        _sut_A._RunExecutionSubstitute();
        _sut_N._RunExecutionSubstitute();
        _done := TRUE;
        ProbeDoneWhen(_done);
    {endregion}
    {region "T505_OnStateChangeWithRestoreCallInside"}
    eTcoSequenceTests.OnStateChangeWithRestoreCallInside:
        IF NOT _arranged THEN
            _sut_A.SetCyclicMode(); //Set sequencer into the cyclic mode
            _sut_N.SetCyclicMode(); //Set sequencer into the cyclic mode
            _sut_A.SetSequenceAsChecked(); //Set sequence as checked, so no StepID uniqueness is performed on next sequence execution
            _sut_N.SetSequenceAsChecked(); //Set sequence as checked, so no StepID uniqueness is performed on next sequence execution
            _sut_A.SetNumberOfSteps(_totalStepNumber); //Set numberOfSteps to the testing instance
            _sut_N.SetNumberOfSteps(_totalStepNumber); //Set numberOfSteps to the testing instance
            _sut_A.TcoSequencerTest := eTcoSequenceTests.OnStateChangeWithRestoreCallInside;
            _sut_N.TcoSequencerTest := eTcoSequenceTests.OnStateChangeWithRestoreCallInside;
            _sut_A.TotalStepNumber := _totalStepNumber;
            _sut_N.TotalStepNumber := _totalStepNumber;
            _sut_A.FinishStep := FALSE;
            _sut_N.FinishStep := FALSE;
            _plcCycleCounter := 0;
            _arranged := TRUE;
            RETURN;
        END_IF

        IF NOT _done THEN
            IF _plcCycleCounter = 1 THEN
                _sut_A.CallRestoreInOnStateChange := FALSE;
                _sut_N.CallRestoreInOnStateChange := FALSE;
            ELSE
                _sut_A.CallRestoreInOnStateChange := TRUE;
                _sut_N.CallRestoreInOnStateChange := TRUE;
                _sut_A.FinishStep := TRUE;
                _sut_N.FinishStep := TRUE;
            END_IF

            _sut_A._RunExecutionSubstitute();
            _sut_N._RunExecutionSubstitute();
        END_IF

        _done := _plcCycleCounter >= 2;

        IF _done THEN
            _sut_A.CallRestoreInOnStateChange := FALSE;
            _sut_N.CallRestoreInOnStateChange := FALSE;
            ProbeDoneWhen(_done);
        END_IF
    {endregion}
    {region "T506_MinStepId"}
    eTcoSequenceTests.MinStepId:
        IF NOT _arranged THEN
            _sut_A.SetCyclicMode(); //Set sequencer into the cyclic mode
            _sut_N.SetCyclicMode(); //Set sequencer into the cyclic mode
            _sut_A.SetSequenceAsChecked(); //Set sequence as checked, so no StepID uniqueness is performed on next sequence execution
            _sut_N.SetSequenceAsChecked(); //Set sequence as checked, so no StepID uniqueness is performed on next sequence execution
            _sut_A.SetNumberOfSteps(_totalStepNumber); //Set numberOfSteps to the testing instance
            _sut_N.SetNumberOfSteps(_totalStepNumber); //Set numberOfSteps to the testing instance
            _sut_A.TcoSequencerTest := eTcoSequenceTests.MinStepId;
            _sut_N.TcoSequencerTest := eTcoSequenceTests.MinStepId;
            _sut_A.TotalStepNumber := _totalStepNumber;
            _sut_N.TotalStepNumber := _totalStepNumber;
            _sut_A.FinishStep := FALSE;
            _sut_N.FinishStep := FALSE;
            _plcCycleCounter := 0;
            _arranged := TRUE;
            RETURN;
        END_IF

        IF NOT _done THEN
            _sut_A.StepId := _currentStepId;
            _sut_N.StepId := _currentStepId;
            _sut_A._RunExecutionSubstitute();
            _sut_N._RunExecutionSubstitute();
        END_IF

        _done := TRUE;
        ProbeDoneWhen(_done);
    {endregion}
    {region "T507_MaxStepId"}
    eTcoSequenceTests.MaxStepId:
        IF NOT _arranged THEN
            _sut_A.SetCyclicMode(); //Set sequencer into the cyclic mode
            _sut_N.SetCyclicMode(); //Set sequencer into the cyclic mode
            _sut_A.SetSequenceAsChecked(); //Set sequence as checked, so no StepID uniqueness is performed on next sequence execution
            _sut_N.SetSequenceAsChecked(); //Set sequence as checked, so no StepID uniqueness is performed on next sequence execution
            _sut_A.SetNumberOfSteps(_totalStepNumber); //Set numberOfSteps to the testing instance
            _sut_N.SetNumberOfSteps(_totalStepNumber); //Set numberOfSteps to the testing instance
            _sut_A.TcoSequencerTest := eTcoSequenceTests.MaxStepId;
            _sut_N.TcoSequencerTest := eTcoSequenceTests.MaxStepId;
            _sut_A.TotalStepNumber := _totalStepNumber;
            _sut_N.TotalStepNumber := _totalStepNumber;
            _sut_A.FinishStep := FALSE;
            _sut_N.FinishStep := FALSE;
            _plcCycleCounter := 0;
            _arranged := TRUE;
            RETURN;
        END_IF

        IF NOT _done THEN
            _sut_A.StepId := _currentStepId;
            _sut_N.StepId := _currentStepId;
            _sut_A._RunExecutionSubstitute();
            _sut_N._RunExecutionSubstitute();
        END_IF

        _done := TRUE;
        ProbeDoneWhen(_done);
    {endregion}
    {region "T508_RequestStepToFirstStepWithStepId0"}
    eTcoSequenceTests.RequestStepToFirstStepWithStepId0:
        IF NOT _arranged THEN
            _sut_A.SetCyclicMode(); //Set sequencer into the cyclic mode
            _sut_N.SetCyclicMode(); //Set sequencer into the cyclic mode
            _sut_A.SetSequenceAsChecked(); //Set sequence as checked, so no StepID uniqueness is performed on next sequence execution
            _sut_N.SetSequenceAsChecked(); //Set sequence as checked, so no StepID uniqueness is performed on next sequence execution
            _sut_A.SetNumberOfSteps(_totalStepNumber); //Set numberOfSteps to the testing instance
            _sut_N.SetNumberOfSteps(_totalStepNumber); //Set numberOfSteps to the testing instance
            _sut_A.TcoSequencerTest := eTcoSequenceTests.RequestStepToFirstStepWithStepId0;
            _sut_N.TcoSequencerTest := eTcoSequenceTests.RequestStepToFirstStepWithStepId0;
            _sut_A.TotalStepNumber := _totalStepNumber;
            _sut_N.TotalStepNumber := _totalStepNumber;
            _sut_A.FinishStep := TRUE;
            _sut_N.FinishStep := TRUE;
            _plcCycleCounter := 0;
            _arranged := TRUE;
            RETURN;
        END_IF

        IF NOT _done THEN
            IF _plcCycleCounter > 1 THEN
                _sut_A.FinishStep := FALSE;
                _sut_N.FinishStep := FalsE;
            END_IF

            _sut_A._RunExecutionSubstitute();
            _sut_N._RunExecutionSubstitute();
        END_IF

        _done := _plcCycleCounter > 1;
        ProbeDoneWhen(_done);
    {endregion}
    {region "T509_RequestStep"}
    eTcoSequenceTests.RequestStep:
        IF NOT _arranged THEN
            _sut_A.SetCyclicMode(); //Set sequencer into the cyclic mode
            _sut_N.SetCyclicMode(); //Set sequencer into the cyclic mode
            _sut_A.SetSequenceAsChecked(); //Set sequence as checked, so no StepID uniqueness is performed on next sequence execution
            _sut_N.SetSequenceAsChecked(); //Set sequence as checked, so no StepID uniqueness is performed on next sequence execution
            _sut_A.SetNumberOfSteps(10); //Set numberOfSteps to the testing instance
            _sut_N.SetNumberOfSteps(10); //Set numberOfSteps to the testing instance
            _sut_A.TcoSequencerTest := eTcoSequenceTests.RequestStep;
            _sut_N.TcoSequencerTest := eTcoSequenceTests.RequestStep;
            _plcCycleCounter := 0;
            _arranged := TRUE;
            RETURN;
        END_IF

        IF NOT _done THEN
            _sut_A.SequenceRun := _plcCycleCounter;
            _sut_N.SequenceRun := _plcCycleCounter;
            _sut_A._RunExecutionSubstitute();
            _sut_N._RunExecutionSubstitute();
        END_IF

        _done := _plcCycleCounter >= 3;
        ProbeDoneWhen(_done);
    {endregion}
    {region "T510_CheckStepIdUniqueness"}
    eTcoSequenceTests.CheckStepIdUniqueness:
        IF NOT _arranged THEN
            _sut_A.SetCyclicMode(); //Set sequencer into the cyclic mode
            _sut_N.SetCyclicMode(); //Set sequencer into the cyclic mode
            _sut_A.SetSequenceAsNotChecked(); //Set sequence as not checked, so StepId uniqueness is going to be performed on next sequence run
            _sut_N.SetSequenceAsNotChecked(); //Set sequence as not checked, so StepId uniqueness is going to be performed on next sequence run
            _sut_A.ClearNumberOfSteps(); //Clear internal step counters, so number of steps is going to be counted again on next sequence run
            _sut_N.ClearNumberOfSteps(); //Clear internal step counters, so number of steps is going to be counted again on next sequence run
            _sut_A.Enabled := TRUE;
            _sut_A.RunOneStep := FALSE;
            _sut_A.RunAllSteps := TRUE;
            _sut_A.FinishStep := TRUE;
            _sut_N.Enabled := TRUE;
            _sut_N.RunOneStep := FALSE;
            _sut_N.RunAllSteps := TRUE;
            _sut_N.FinishStep := TRUE;
            _sut_A.SetCurrentStep(inStepID := _currentStepId, inStepDescription := _currentStepDescription);
            _sut_N.SetCurrentStep(inStepID := _currentStepId, inStepDescription := _currentStepDescription);
            _sut_A.TcoSequencerTest := eTcoSequenceTests.CheckStepIdUniqueness;
            _sut_N.TcoSequencerTest := eTcoSequenceTests.CheckStepIdUniqueness;
            _sut_A.SaveNumberOfStepsInSequence();
            _sut_N.SaveNumberOfStepsInSequence();
            _plcCycleCounter := 0;
            _arranged := TRUE;
            RETURN;
        END_IF

        IF NOT _done THEN
            _sut_A._RunExecutionSubstitute();
            _sut_N._RunExecutionSubstitute();
            _sut_A.SaveNumberOfStepsInSequence();
            _sut_N.SaveNumberOfStepsInSequence();
        END_IF

        _done := _plcCycleCounter >= 2;
        ProbeDoneWhen(_done);
    {endregion}
    {region "T512_RestoreAlreadyCheckedSequence"}
    eTcoSequenceTests.RestoreAlreadyCheckedSequence:
        _sut_A.Restore();
        _sut_N.Restore();
        _sut_A.SaveNumberOfStepsInSequence();
        _sut_N.SaveNumberOfStepsInSequence();
        _done := TRUE;
        ProbeDoneWhen(_done);
    {endregion}
    {region "T513_CheckStepIdUniqueness"}
    eTcoSequenceTests.NotUniqueStepId:
        IF NOT _arranged THEN
            _sut_A.Enabled := TRUE;
            _sut_A.RunOneStep := FALSE;
            _sut_A.RunAllSteps := FALSE;
            _sut_A.FinishStep := TRUE;
            _sut_A.StepId := _stepId;
            _sut_N.Enabled := TRUE;
            _sut_N.RunOneStep := FALSE;
            _sut_N.RunAllSteps := FALSE;
            _sut_N.FinishStep := TRUE;
            _sut_N.StepId := _stepId;
            _sut_A.SetCurrentStep(inStepID := _currentStepId, inStepDescription := _currentStepDescription);
            _sut_N.SetCurrentStep(inStepID := _currentStepId, inStepDescription := _currentStepDescription);
            _sut_A.TcoSequencerTest := eTcoSequenceTests.NotUniqueStepId;
            _sut_N.TcoSequencerTest := eTcoSequenceTests.NotUniqueStepId;
            _sut_A.SaveNumberOfStepsInSequence();
            _sut_N.SaveNumberOfStepsInSequence();
            _plcCycleCounter := 0;
			_sut_A._messenger.Clear();
			_sut_N._messenger.Clear();
            _arranged := TRUE;
            RETURN;
        END_IF

        IF NOT _done THEN								 
            _sut_A._RunExecutionSubstitute();
            _sut_N._RunExecutionSubstitute();
            _sut_A.SaveNumberOfStepsInSequence();
            _sut_N.SaveNumberOfStepsInSequence();
            _done := _plcCycleCounter >= 2;
        END_IF

        IF _done THEN
            ProbeDoneWhen(_done);
        END_IF
    {endregion}
    {region "T516_AfterErrorRestore"}
    eTcoSequenceTests.AfterErrorRestore:
        IF NOT _arranged THEN
            _sut_A.TcoSequencerTest := eTcoSequenceTests.AfterErrorRestore;
            _sut_N.TcoSequencerTest := eTcoSequenceTests.AfterErrorRestore;
            _sut_A.SaveNumberOfStepsInSequence();
            _sut_N.SaveNumberOfStepsInSequence();
            _plcCycleCounter := 0;
            _arranged := TRUE;
            RETURN;
        END_IF

        IF NOT _done THEN
            _sut_A._RunExecutionSubstitute();
            _sut_N._RunExecutionSubstitute();
            _sut_A.SaveNumberOfStepsInSequence();
            _sut_N.SaveNumberOfStepsInSequence();
            _done := _plcCycleCounter >= 3;
        END_IF

        IF _done THEN
            ProbeDoneWhen(_done);
        END_IF
    {endregion}
    {region "T520_ChangeStepIdDuringExecution"}
    eTcoSequenceTests.ChangeStepIdDuringExecution:
        IF NOT _arranged THEN
            _sut_A.TcoSequencerTest := eTcoSequenceTests.ChangeStepIdDuringExecution;
            _sut_N.TcoSequencerTest := eTcoSequenceTests.ChangeStepIdDuringExecution;
            _sut_A.SetCyclicMode(); //Set sequencer into the cyclic mode
            _sut_N.SetCyclicMode(); //Set sequencer into the cyclic mode
            _sut_A.SetSequenceAsChecked(); //Set sequence as checked, so no StepID uniqueness is performed on next sequence execution
            _sut_N.SetSequenceAsChecked(); //Set sequence as checked, so no StepID uniqueness is performed on next sequence execution
            _sut_A.ClearNumberOfSteps(); //Clear internal step counters, so number of steps is going to be counted again on next sequence run
            _sut_N.ClearNumberOfSteps(); //Clear internal step counters, so number of steps is going to be counted again on next sequence run
            _sut_A.SetCurrentStep(inStepID := _currentStepId, inStepDescription := _currentStepDescription);
            _sut_N.SetCurrentStep(inStepID := _currentStepId, inStepDescription := _currentStepDescription);
            _sut_A.TotalStepNumber := _totalStepNumber;
            _sut_N.TotalStepNumber := _totalStepNumber;
            _sut_A.SaveNumberOfStepsInSequence();
            _sut_N.SaveNumberOfStepsInSequence();
            _plcCycleCounter := 0;
            _arranged := TRUE;
            RETURN;
        END_IF

        IF NOT _done THEN
            _sut_A.SequenceRun := _plcCycleCounter;
            _sut_N.SequenceRun := _plcCycleCounter;
            _sut_A._RunExecutionSubstitute();
            _sut_N._RunExecutionSubstitute();
            _sut_A.SaveNumberOfStepsInSequence();
            _sut_N.SaveNumberOfStepsInSequence();
        END_IF

        _done := _plcCycleCounter >= 3;
        ProbeDoneWhen(_done);
    {endregion}
    {region "T524_CommentOutPartOfRunningSequencer"}
    eTcoSequenceTests.CommentOutPartOfRunningSequencer:
        IF NOT _arranged THEN
            _sut_A.TcoSequencerTest := eTcoSequenceTests.CommentOutPartOfRunningSequencer;
            _sut_N.TcoSequencerTest := eTcoSequenceTests.CommentOutPartOfRunningSequencer;
            _sut_A.SetCyclicMode(); //Set sequencer into the cyclic mode
            _sut_N.SetCyclicMode(); //Set sequencer into the cyclic mode
            _sut_A.SetSequenceAsChecked(); //Set sequence as checked, so no StepID uniqueness is performed on next sequence execution
            _sut_N.SetSequenceAsChecked(); //Set sequence as checked, so no StepID uniqueness is performed on next sequence execution
            _sut_A.ClearNumberOfSteps(); //Clear internal step counters, so number of steps is going to be counted again on next sequence run
            _sut_N.ClearNumberOfSteps(); //Clear internal step counters, so number of steps is going to be counted again on next sequence run
            _sut_A.SetCurrentStep(inStepID := _currentStepId, inStepDescription := _currentStepDescription);
            _sut_N.SetCurrentStep(inStepID := _currentStepId, inStepDescription := _currentStepDescription);
            _sut_A.TotalStepNumber := _totalStepNumber;
            _sut_N.TotalStepNumber := _totalStepNumber;
            _sut_A.SaveNumberOfStepsInSequence();
            _sut_N.SaveNumberOfStepsInSequence();
            _plcCycleCounter := 0;
            _arranged := TRUE;
            RETURN;
        END_IF

        IF NOT _done THEN
            IF _plcCycleCounter = 3 THEN
                _sut_A.Restore();
                _sut_N.Restore();
                _sut_A.SetSequenceAsChecked(); //Set sequence as checked, so no StepID uniqueness is performed on next sequence execution
                _sut_N.SetSequenceAsChecked(); //Set sequence as checked, so no StepID uniqueness is performed on next sequence execution
                _sut_A.ClearNumberOfSteps(); //Clear internal step counters, so number of steps is going to be counted again on next sequence run
                _sut_N.ClearNumberOfSteps(); //Clear internal step counters, so number of steps is going to be counted again on next sequence run
            END_IF

            _sut_A.SequenceRun := _plcCycleCounter;
            _sut_N.SequenceRun := _plcCycleCounter;
            _sut_A._RunExecutionSubstitute();
            _sut_N._RunExecutionSubstitute();
            _sut_A.SaveNumberOfStepsInSequence();
            _sut_N.SaveNumberOfStepsInSequence();
        END_IF

        _done := _plcCycleCounter >= 3;
        ProbeDoneWhen(_done);
    {endregion}
    {region "T526_UncommentPartOfRunningSequencer"}
    eTcoSequenceTests.UncommentPartOfRunningSequencer:
        IF NOT _arranged THEN
            _sut_A.TcoSequencerTest := eTcoSequenceTests.UncommentPartOfRunningSequencer;
            _sut_N.TcoSequencerTest := eTcoSequenceTests.UncommentPartOfRunningSequencer;
            _sut_A.SetCyclicMode(); //Set sequencer into the cyclic mode
            _sut_N.SetCyclicMode(); //Set sequencer into the cyclic mode
            _sut_A.SetSequenceAsChecked(); //Set sequence as checked, so no StepID uniqueness is performed on next sequence execution
            _sut_N.SetSequenceAsChecked(); //Set sequence as checked, so no StepID uniqueness is performed on next sequence execution
            _sut_A.ClearNumberOfSteps(); //Clear internal step counters, so number of steps is going to be counted again on next sequence run
            _sut_N.ClearNumberOfSteps(); //Clear internal step counters, so number of steps is going to be counted again on next sequence run
            _sut_A.SetCurrentStep(inStepID := _currentStepId, inStepDescription := _currentStepDescription);
            _sut_N.SetCurrentStep(inStepID := _currentStepId, inStepDescription := _currentStepDescription);
            _sut_A.TotalStepNumber := _totalStepNumber;
            _sut_N.TotalStepNumber := _totalStepNumber;
            _sut_A.SaveNumberOfStepsInSequence();
            _sut_N.SaveNumberOfStepsInSequence();
            _plcCycleCounter := 0;
            _arranged := TRUE;
            RETURN;
        END_IF

        IF NOT _done THEN
            _sut_A.SequenceRun := _plcCycleCounter;
            _sut_N.SequenceRun := _plcCycleCounter;
            _sut_A._RunExecutionSubstitute();
            _sut_N._RunExecutionSubstitute();
            _sut_A.SaveNumberOfStepsInSequence();
            _sut_N.SaveNumberOfStepsInSequence();
        END_IF

        _done := _plcCycleCounter >= 2;
        ProbeDoneWhen(_done);
    {endregion}
    {region "T530_OpenCloseSequence"}
    eTcoSequenceTests.OpenCloseSequence:
        IF NOT _arranged THEN
            _sut_A.TcoSequencerTest := eTcoSequenceTests.OpenCloseSequence;
            _sut_N.TcoSequencerTest := eTcoSequenceTests.OpenCloseSequence;
            _sut_A.SetCyclicMode(); //Set sequencer into the cyclic mode
            _sut_N.SetCyclicMode(); //Set sequencer into the cyclic mode
            _sut_A.SetSequenceAsChecked(); //Set sequence as checked, so no StepID uniqueness is performed on next sequence execution
            _sut_N.SetSequenceAsChecked(); //Set sequence as checked, so no StepID uniqueness is performed on next sequence execution
            _sut_A.ClearNumberOfSteps(); //Clear internal step counters, so number of steps is going to be counted again on next sequence run
            _sut_N.ClearNumberOfSteps(); //Clear internal step counters, so number of steps is going to be counted again on next sequence run
            _sut_A.TotalStepNumber := _totalStepNumber;
            _sut_N.TotalStepNumber := _totalStepNumber;
            _sut_A.SaveNumberOfStepsInSequence();
            _sut_N.SaveNumberOfStepsInSequence();
            _plcCycleCounter := 0;
            _arranged := TRUE;
            RETURN;
        END_IF

        IF NOT _done THEN
            IF _plcCycleCounter = 1 THEN
                _sut_A.SequencerOpen();
                _sut_N.SequencerOpen();

                IF _sut_A._Step(0, TRUE, 'Step 0') THEN
                    _sut_A._StepCompleteWhen(TRUE);
                END_IF

                IF _sut_N._Step(0, TRUE, 'Step 0') THEN
                    _sut_N._StepCompleteWhen(TRUE);
                END_IF
				_sut_A.SequencerClose();
                _sut_N.SequencerClose();
            END_IF

            IF _plcCycleCounter = 2 THEN
				_sut_A.SequencerOpen();
                _sut_N.SequencerOpen();
                FOR i := 1 TO _totalStepNumber DO
                    _sut_A._Step(i, TRUE, CONCAT('Step ', INT_TO_STRING(i)));
                    _sut_N._Step(i, TRUE, CONCAT('Step ', INT_TO_STRING(i)));
                END_FOR

                _sut_A.SequencerClose();
                _sut_N.SequencerClose();
            END_IF
		END_IF;		 
		
        _done := _plcCycleCounter >= 2;
        ProbeDoneWhen(_done);			  

//            IF _plcCycleCounter = 3 THEN
//                _sut_A.SequencerOpen();
//                _sut_N.SequencerOpen();
//			    _sut_A.SequencerClose();
//                _sut_N.SequencerClose();
//            END_IF

//            IF _plcCycleCounter = 4 THEN
//				_sut_A.SequencerOpen();
//                _sut_N.SequencerOpen();
//                IF _sut_A._Step(0, TRUE, 'Step 0') THEN
//                    _sut_A._StepCompleteWhen(TRUE);
//                END_IF

//                IF _sut_N._Step(0, TRUE, 'Step 0') THEN
//                    _sut_N._StepCompleteWhen(TRUE);
//                END_IF
//				_sut_A.SequencerClose();
//                _sut_N.SequencerClose();	 
//            END_IF

//            IF _plcCycleCounter = 5 THEN
//				_sut_A.SequencerOpen();
//                _sut_N.SequencerOpen();
//                FOR i := 1 TO _totalStepNumber DO
//                    IF _sut_A._Step(i, TRUE, CONCAT('Step ', INT_TO_STRING(i))) THEN
//                        _sut_A._StepCompleteWhen(TRUE);
//                    END_IF

//                    IF _sut_N._Step(i, TRUE, CONCAT('Step ', INT_TO_STRING(i))) THEN
//                        _sut_N._StepCompleteWhen(TRUE);
//                    END_IF
//                END_FOR
//				_sut_A.SequencerClose();
//                _sut_N.SequencerClose();	 
//            END_IF

//            IF _plcCycleCounter = 6 THEN
//                _sut_A._SequenceComplete();
//                _sut_N._SequenceComplete();
//                _sut_A.SequencerClose();
//                _sut_N.SequencerClose();
//            END_IF

//            IF _plcCycleCounter = 7 THEN
//                _sut_A.SequencerOpen();
//                _sut_N.SequencerOpen();
//            END_IF

//            IF _plcCycleCounter = 8 THEN
//                _sut_A.SequencerClose();
//                _sut_N.SequencerClose();
//            END_IF

//            IF _plcCycleCounter = 9 THEN
//                _sut_A.SequencerOpen();
//                _sut_N.SequencerOpen();
//                _sut_A._Step(0, TRUE, 'Step 0');
//                _sut_N._Step(0, TRUE, 'Step 0');
//                _sut_A.SequencerClose();
//                _sut_N.SequencerClose();
//            END_IF
//        END_IF

//        _done := _plcCycleCounter >= 9;
//        ProbeDoneWhen(_done);
    {endregion}
    {region "T541_RequestStepFromLowerToHigher"}
    eTcoSequenceTests.RequestStepFromLowerToHigher:
        IF NOT _arranged THEN
            _sut_A.TcoSequencerTest := eTcoSequenceTests.RequestStepFromLowerToHigher;
            _sut_N.TcoSequencerTest := eTcoSequenceTests.RequestStepFromLowerToHigher;
            _sut_A.SetCyclicMode(); //Set sequencer into the cyclic mode
            _sut_N.SetCyclicMode(); //Set sequencer into the cyclic mode
            _sut_A.SetSequenceAsChecked(); //Set sequence as checked, so no StepID uniqueness is performed on next sequence execution
            _sut_N.SetSequenceAsChecked(); //Set sequence as checked, so no StepID uniqueness is performed on next sequence execution
            _sut_A.ClearNumberOfSteps(); //Clear internal step counters, so number of steps is going to be counted again on next sequence run
            _sut_N.ClearNumberOfSteps(); //Clear internal step counters, so number of steps is going to be counted again on next sequence run
            _sut_A.SetCurrentStep(inStepID := _currentStepId, inStepDescription := _currentStepDescription);
            _sut_N.SetCurrentStep(inStepID := _currentStepId, inStepDescription := _currentStepDescription);
            _sut_A.TotalStepNumber := _totalStepNumber;
            _sut_N.TotalStepNumber := _totalStepNumber;
            _sut_A.ReqStep := _reqStep;
            _sut_N.ReqStep := _reqStep;
            _sut_A.ReqStepNotExists := _reqStepNotExists;
            _sut_N.ReqStepNotExists := _reqStepNotExists;
            _sut_A.SaveNumberOfStepsInSequence();
            _sut_N.SaveNumberOfStepsInSequence();
            _plcCycleCounter := 0;
            _arranged := TRUE;
            RETURN;
        END_IF

        IF NOT _done THEN
            _sut_A.SequenceRun := _plcCycleCounter;
            _sut_N.SequenceRun := _plcCycleCounter;
            _sut_A._RunExecutionSubstitute();
            _sut_N._RunExecutionSubstitute();
            _sut_A.SaveNumberOfStepsInSequence();
            _sut_N.SaveNumberOfStepsInSequence();
        END_IF

        _done := _plcCycleCounter >= 2;
        ProbeDoneWhen(_done);
    {endregion}
    {region "T542_RequestStepFromHigherToLower"}
    eTcoSequenceTests.RequestStepFromHigherToLower:
        IF NOT _arranged THEN
            _sut_A.TcoSequencerTest := eTcoSequenceTests.RequestStepFromHigherToLower;
            _sut_N.TcoSequencerTest := eTcoSequenceTests.RequestStepFromHigherToLower;
            _sut_A.SetCyclicMode(); //Set sequencer into the cyclic mode
            _sut_N.SetCyclicMode(); //Set sequencer into the cyclic mode
            _sut_A.SetSequenceAsChecked(); //Set sequence as checked, so no StepID uniqueness is performed on next sequence execution
            _sut_N.SetSequenceAsChecked(); //Set sequence as checked, so no StepID uniqueness is performed on next sequence execution
            _sut_A.SetNumberOfSteps(_totalStepNumber);
            _sut_N.SetNumberOfSteps(_totalStepNumber);
            _sut_A.SetCurrentStep(inStepID := _currentStepId, inStepDescription := _currentStepDescription);
            _sut_N.SetCurrentStep(inStepID := _currentStepId, inStepDescription := _currentStepDescription);
            _sut_A.TotalStepNumber := _totalStepNumber;
            _sut_N.TotalStepNumber := _totalStepNumber;
            _sut_A.ReqStep := _reqStep;
            _sut_N.ReqStep := _reqStep;
            _sut_A.ReqStepNotExists := _reqStepNotExists;
            _sut_N.ReqStepNotExists := _reqStepNotExists;
            _sut_A.SaveNumberOfStepsInSequence();
            _sut_N.SaveNumberOfStepsInSequence();
            _plcCycleCounter := 0;
            _arranged := TRUE;
            RETURN;
        END_IF

        IF NOT _done THEN
            _sut_A.SequenceRun := _plcCycleCounter;
            _sut_N.SequenceRun := _plcCycleCounter;
            _sut_A._RunExecutionSubstitute();
            _sut_N._RunExecutionSubstitute();
            _sut_A.SaveNumberOfStepsInSequence();
            _sut_N.SaveNumberOfStepsInSequence();
        END_IF

        _done := _plcCycleCounter >= 2;
        ProbeDoneWhen(_done);
    {endregion}
    {region "T544_RequestStepToNotExistingStep"}
    eTcoSequenceTests.RequestStepToNotExistingStep:
        IF NOT _arranged THEN
            _sut_A.TcoSequencerTest := eTcoSequenceTests.RequestStepToNotExistingStep;
            _sut_N.TcoSequencerTest := eTcoSequenceTests.RequestStepToNotExistingStep;
            _sut_A.SetCyclicMode(); //Set sequencer into the cyclic mode
            _sut_N.SetCyclicMode(); //Set sequencer into the cyclic mode
            _sut_A.SetSequenceAsChecked(); //Set sequence as checked, so no StepID uniqueness is performed on next sequence execution
            _sut_N.SetSequenceAsChecked(); //Set sequence as checked, so no StepID uniqueness is performed on next sequence execution
            _sut_A.SetNumberOfSteps(_totalStepNumber);
            _sut_N.SetNumberOfSteps(_totalStepNumber);
            _sut_A.SetCurrentStep(inStepID := _currentStepId, inStepDescription := _currentStepDescription);
            _sut_N.SetCurrentStep(inStepID := _currentStepId, inStepDescription := _currentStepDescription);
            _sut_A.TotalStepNumber := _totalStepNumber;
            _sut_N.TotalStepNumber := _totalStepNumber;
            _sut_A.ReqStep := _reqStep;
            _sut_N.ReqStep := _reqStep;
            _sut_A.ReqStepNotExists := _reqStepNotExists;
            _sut_N.ReqStepNotExists := _reqStepNotExists;
            _sut_A.SaveNumberOfStepsInSequence();
            _sut_N.SaveNumberOfStepsInSequence();
            _plcCycleCounter := 0;
            _arranged := TRUE;
            RETURN;
        END_IF

        IF _plcCycleCounter = 4 THEN
            _sut_A.Restore();
            _sut_N.Restore();
            _sut_A.SetCyclicMode(); //Set sequencer into the cyclic mode
            _sut_N.SetCyclicMode(); //Set sequencer into the cyclic mode
            _sut_A.SetSequenceAsChecked(); //Set sequence as checked, so no StepID uniqueness is performed on next sequence execution
            _sut_N.SetSequenceAsChecked(); //Set sequence as checked, so no StepID uniqueness is performed on next sequence execution
            _sut_A.SetNumberOfSteps(_totalStepNumber);
            _sut_N.SetNumberOfSteps(_totalStepNumber);
            _sut_A.SetCurrentStep(inStepID := _currentStepId, inStepDescription := _currentStepDescription);
            _sut_N.SetCurrentStep(inStepID := _currentStepId, inStepDescription := _currentStepDescription);
            _sut_A.TotalStepNumber := _totalStepNumber;
            _sut_N.TotalStepNumber := _totalStepNumber;
        END_IF

        IF NOT _done THEN
            _sut_A.SequenceRun := _plcCycleCounter;
            _sut_N.SequenceRun := _plcCycleCounter;
            _sut_A._RunExecutionSubstitute();
            _sut_N._RunExecutionSubstitute();
            _sut_A.SaveNumberOfStepsInSequence();
            _sut_N.SaveNumberOfStepsInSequence();
        END_IF

        _done := _plcCycleCounter >= 4;
        ProbeDoneWhen(_done);
    {endregion}
    {region "T547_RequestStepWhilePreviousRequestStepHasNotBeenYetProcessed"}
    eTcoSequenceTests.RequestStepWhilePreviousRequestStepHasNotBeenYetProcessed:
        IF NOT _arranged THEN
            _sut_A.TcoSequencerTest := eTcoSequenceTests.RequestStepWhilePreviousRequestStepHasNotBeenYetProcessed;
            _sut_N.TcoSequencerTest := eTcoSequenceTests.RequestStepWhilePreviousRequestStepHasNotBeenYetProcessed;
            _sut_A.SetCyclicMode(); //Set sequencer into the cyclic mode
            _sut_N.SetCyclicMode(); //Set sequencer into the cyclic mode
            _sut_A.SetSequenceAsChecked(); //Set sequence as checked, so no StepID uniqueness is performed on next sequence execution
            _sut_N.SetSequenceAsChecked(); //Set sequence as checked, so no StepID uniqueness is performed on next sequence execution
            _sut_A.SetNumberOfSteps(_totalStepNumber);
            _sut_N.SetNumberOfSteps(_totalStepNumber);
            _sut_A.SetCurrentStep(inStepID := _currentStepId, inStepDescription := _currentStepDescription);
            _sut_N.SetCurrentStep(inStepID := _currentStepId, inStepDescription := _currentStepDescription);
            _sut_A.TotalStepNumber := _totalStepNumber;
            _sut_N.TotalStepNumber := _totalStepNumber;
            _sut_A.ReqStep := _reqStep;
            _sut_N.ReqStep := _reqStep;
            _sut_A.ReqStepNotExists := _reqStepNotExists;
            _sut_N.ReqStepNotExists := _reqStepNotExists;
            _sut_A.SaveNumberOfStepsInSequence();
            _sut_N.SaveNumberOfStepsInSequence();
            _plcCycleCounter := 0;
            _arranged := TRUE;
            RETURN;
        END_IF

        IF NOT _done THEN
            _sut_A.SequenceRun := _plcCycleCounter;
            _sut_N.SequenceRun := _plcCycleCounter;
            _sut_A._RunExecutionSubstitute();
            _sut_N._RunExecutionSubstitute();
            _sut_A.SaveNumberOfStepsInSequence();
            _sut_N.SaveNumberOfStepsInSequence();
        END_IF

        _done := TRUE;
        ProbeDoneWhen(_done);
    {endregion}
    {region "T551_DisableStepEnabledAndActiveInPreviousPLCcycle"}
    eTcoSequenceTests.DisableStepEnabledAndActiveInPreviousPLCcycle:
        IF NOT _arranged THEN
            _sut_A.TcoSequencerTest := eTcoSequenceTests.DisableStepEnabledAndActiveInPreviousPLCcycle;
            _sut_N.TcoSequencerTest := eTcoSequenceTests.DisableStepEnabledAndActiveInPreviousPLCcycle;
            _sut_A.SetCyclicMode(); //Set sequencer into the cyclic mode
            _sut_N.SetCyclicMode(); //Set sequencer into the cyclic mode
            _sut_A.SetSequenceAsChecked(); //Set sequence as checked, so no StepID uniqueness is performed on next sequence execution
            _sut_N.SetSequenceAsChecked(); //Set sequence as checked, so no StepID uniqueness is performed on next sequence execution
            _sut_A.SetNumberOfSteps(_totalStepNumber);
            _sut_N.SetNumberOfSteps(_totalStepNumber);
            _sut_A.TotalStepNumber := _totalStepNumber;
            _sut_N.TotalStepNumber := _totalStepNumber;
            _sut_A.SaveNumberOfStepsInSequence();
            _sut_N.SaveNumberOfStepsInSequence();
            _plcCycleCounter := 0;
            _arranged := TRUE;
            RETURN;
        END_IF

        IF NOT _done THEN
            IF _plcCycleCounter = 1 THEN
                _sut_A.SequencerOpen();

                IF _sut_A._Step(0, TRUE, 'Step 0') THEN
                    _sut_A._StepCompleteWhen(TRUE);
                END_IF

                FOR i := 1 TO _totalStepNumber - 2 DO
                    _sut_A._Step(i, TRUE, CONCAT('Step ', INT_TO_STRING(i)));
                END_FOR

                IF _sut_A._Step(_totalStepNumber - 1, TRUE, CONCAT('Step ', INT_TO_STRING(_totalStepNumber - 1))) THEN
                    _sut_A._SequenceComplete();
                END_IF

                _sut_A.SequencerClose();
                _sut_N.SequencerOpen();

                IF _sut_N._Step(0, TRUE, 'Step 0') THEN
                    _sut_N._StepCompleteWhen(TRUE);
                END_IF

                FOR i := 1 TO _totalStepNumber - 2 DO
                    _sut_N._Step(i, TRUE, CONCAT('Step ', INT_TO_STRING(i)));
                END_FOR

                IF _sut_N._Step(_totalStepNumber - 1, TRUE, CONCAT('Step ', INT_TO_STRING(_totalStepNumber - 1))) THEN
                    _sut_N._SequenceComplete();
                END_IF

                _sut_N.SequencerClose();
            END_IF

            IF _plcCycleCounter = 2 THEN
                _sut_A.SequencerOpen();

                IF _sut_A._Step(0, TRUE, 'Step 0') THEN
                    _sut_A._StepCompleteWhen(TRUE);
                END_IF

                IF _sut_A._Step(1, FALSE, 'Step 0') THEN
                    _sut_A._StepCompleteWhen(FALSE);
                END_IF

                _sut_N.SequencerOpen();

                IF _sut_N._Step(0, TRUE, 'Step 0') THEN
                    _sut_N._StepCompleteWhen(TRUE);
                END_IF

                IF _sut_N._Step(1, FALSE, 'Step 0') THEN
                    _sut_N._StepCompleteWhen(FALSE);
                END_IF
            END_IF

            IF _plcCycleCounter = 3 THEN
                FOR i := 2 TO _totalStepNumber - 2 DO
                    _sut_A._Step(i, TRUE, CONCAT('Step ', INT_TO_STRING(i)));
                END_FOR

                IF _sut_A._Step(_totalStepNumber - 1, TRUE, CONCAT('Step ', INT_TO_STRING(_totalStepNumber - 1))) THEN
                    _sut_A._SequenceComplete();
                END_IF

                _sut_A.SequencerClose();

                FOR i := 2 TO _totalStepNumber - 2 DO
                    _sut_N._Step(i, TRUE, CONCAT('Step ', INT_TO_STRING(i)));
                END_FOR

                IF _sut_N._Step(_totalStepNumber - 1, TRUE, CONCAT('Step ', INT_TO_STRING(_totalStepNumber - 1))) THEN
                    _sut_N._SequenceComplete();
                END_IF

                _sut_N.SequencerClose();
            END_IF

            _sut_A.SaveNumberOfStepsInSequence();
            _sut_N.SaveNumberOfStepsInSequence();
        END_IF

        _done := _plcCycleCounter >= 3;
        ProbeDoneWhen(_done);
    {endregion}
    {region "T560_RequestStepCallingCyclically"}
    eTcoSequenceTests.RequestStepCallingCyclically:
        IF NOT _arranged THEN
            _sut_A.TcoSequencerTest := eTcoSequenceTests.RequestStepCallingCyclically;
            _sut_N.TcoSequencerTest := eTcoSequenceTests.RequestStepCallingCyclically;
            _sut_A.SetCyclicMode(); //Set sequencer into the cyclic mode
            _sut_N.SetCyclicMode(); //Set sequencer into the cyclic mode
            _sut_A.SetSequenceAsChecked(); //Set sequence as checked, so no StepID uniqueness is performed on next sequence execution
            _sut_N.SetSequenceAsChecked(); //Set sequence as checked, so no StepID uniqueness is performed on next sequence execution
            _sut_A.SetNumberOfSteps(_totalStepNumber);
            _sut_N.SetNumberOfSteps(_totalStepNumber);
            _sut_A.TotalStepNumber := _totalStepNumber;
            _sut_N.TotalStepNumber := _totalStepNumber;
            _sut_A.InitReqStepCycle := _initReqStepCycle;
            _sut_N.InitReqStepCycle := _initReqStepCycle;
            _sut_A.SaveNumberOfStepsInSequence();
            _sut_N.SaveNumberOfStepsInSequence();
            _plcCycleCounter := 0;
            _arranged := TRUE;
            RETURN;
        END_IF

        IF NOT _done THEN
            IF _plcCycleCounter = 1 THEN
                _sut_A.SequencerOpen();
                _sut_N.SequencerOpen();
            END_IF

            IF _plcCycleCounter = 2 THEN
                _sut_A.SequencerOpen();
                _sut_A._RequestStep(10);
                _sut_A.SequencerClose();
                _sut_A.SequencerOpen();
                _sut_N.SequencerOpen();
                _sut_N._RequestStep(10);
                _sut_N.SequencerClose();
                _sut_N.SequencerOpen();
            END_IF

            IF _plcCycleCounter = 3 THEN
                _sut_A._Step(0, TRUE, 'Step 0');
                _sut_A._Step(20, TRUE, 'Step 20');
                _sut_A._Step(10, TRUE, 'Step 10');
                _sut_A.SequencerClose();
                _sut_N._Step(0, TRUE, 'Step 0');
                _sut_N._Step(20, TRUE, 'Step 20');
                _sut_N._Step(10, TRUE, 'Step 10');
                _sut_N.SequencerClose();
            END_IF

            IF _plcCycleCounter = 4 THEN
                _sut_A.InitReqStepCycle := _initReqStepCycle;
                _sut_N.InitReqStepCycle := _initReqStepCycle;
            END_IF

            IF _plcCycleCounter >= 5 THEN
                _sut_A.SequencerOpen();
                _sut_A.PostOpenRequestStepCycle := _sut_A.RequestStepCycle;
                _sut_A._Step(0, TRUE, 'Step 0');

                IF (_sut_A._Step(20, TRUE, 'Step 20')) THEN
                    _sut_A._RequestStep(20);
                END_IF

                IF (_sut_A._Step(10, TRUE, 'Step 10')) THEN
                    _sut_A._RequestStep(20);
                END_IF

                _sut_A.PreCloseRequestStepCycle := _sut_A.RequestStepCycle;
                _sut_A.SequencerClose();
                _sut_N.SequencerOpen();
                _sut_N.PostOpenRequestStepCycle := _sut_N.RequestStepCycle;
                _sut_N._Step(0, TRUE, 'Step 0');

                IF (_sut_N._Step(20, TRUE, 'Step 20')) THEN
                    _sut_N._RequestStep(20);
                END_IF

                IF (_sut_N._Step(10, TRUE, 'Step 10')) THEN
                    _sut_N._RequestStep(20);
                END_IF

                _sut_N.PreCloseRequestStepCycle := _sut_N.RequestStepCycle;
                _sut_N.SequencerClose();
            END_IF
        END_IF

        _sut_A.SaveNumberOfStepsInSequence();
        _sut_N.SaveNumberOfStepsInSequence();
        _done := _plcCycleCounter >= _cycles + 4;
        ProbeDoneWhen(_done);
    {endregion}
    {region "T570_SetStepMode"}
    eTcoSequenceTests.SetStepMode:
        IF NOT _arranged THEN
            _sut_A.TcoSequencerTest := eTcoSequenceTests.SetStepMode;
            _sut_N.TcoSequencerTest := eTcoSequenceTests.SetStepMode;
            _sut_A.SetStepMode(); //Set sequencer into the step mode
            _sut_N.SetStepMode(); //Set sequencer into the step mode
            _sut_A.SetSequenceAsChecked(); //Set sequence as checked, so no StepID uniqueness is performed on next sequence execution
            _sut_N.SetSequenceAsChecked(); //Set sequence as checked, so no StepID uniqueness is performed on next sequence execution
            _sut_A.ClearNumberOfSteps();
            _sut_N.ClearNumberOfSteps();
            _sut_A.SetCurrentStep(inStepID := _currentStepId, inStepDescription := _currentStepDescription);
            _sut_N.SetCurrentStep(inStepID := _currentStepId, inStepDescription := _currentStepDescription);
            _sut_A.TotalStepNumber := _totalStepNumber;
            _sut_N.TotalStepNumber := _totalStepNumber;
            _sut_A.SaveNumberOfStepsInSequence();
            _sut_N.SaveNumberOfStepsInSequence();
            _plcCycleCounter := 0;
            _arranged := TRUE;
            RETURN;
        END_IF

        IF NOT _done THEN
            _sut_A.SequenceRun := _plcCycleCounter;
            _sut_N.SequenceRun := _plcCycleCounter;

            IF _plcCycleCounter = 1 THEN
                _sut_A._RunExecutionSubstitute();
                _sut_N._RunExecutionSubstitute();
            END_IF

            IF _plcCycleCounter = 2 THEN
                _sut_A.SequencerOpen();
                _sut_A._StepIn();

                IF _sut_A._Step(0, TRUE, 'Initial step') THEN
                    _sut_A._StepCompleteWhen(TRUE);
                END_IF

                _sut_N.SequencerOpen();
                _sut_N._StepIn();

                IF _sut_N._Step(0, TRUE, 'Initial step') THEN
                    _sut_N._StepCompleteWhen(TRUE);
                END_IF
            END_IF

            IF _plcCycleCounter = 3 THEN
                IF _sut_A._Step(1, TRUE, 'Step 1') THEN
                    _sut_A._StepCompleteWhen(TRUE);
                END_IF

                IF _sut_N._Step(1, TRUE, 'Step 1') THEN
                    _sut_N._StepCompleteWhen(TRUE);
                END_IF

                FOR i := 2 TO _totalStepNumber - 2 DO
                    _sut_A._Step(i, TRUE, CONCAT('Step ', INT_TO_STRING(i)));
                    _sut_N._Step(i, TRUE, CONCAT('Step ', INT_TO_STRING(i)));
                END_FOR

                IF _sut_A._Step(_totalStepNumber - 1, TRUE, CONCAT('Step ', INT_TO_STRING(_totalStepNumber - 1))) THEN
                    _sut_A._SequenceComplete();
                END_IF

                IF _sut_N._Step(_totalStepNumber - 1, TRUE, CONCAT('Step ', INT_TO_STRING(_totalStepNumber - 1))) THEN
                    _sut_N._SequenceComplete();
                END_IF
            END_IF

            IF _plcCycleCounter = 4 THEN
                _sut_A._RunExecutionSubstitute();
                _sut_N._RunExecutionSubstitute();
            END_IF

            _sut_A.SaveNumberOfStepsInSequence();
            _sut_N.SaveNumberOfStepsInSequence();
        END_IF

        _done := _plcCycleCounter >= 4;
        ProbeDoneWhen(_done);
    {endregion}
    {region "T580_StepMode"}
    eTcoSequenceTests.StepMode:
        IF NOT _arranged THEN
            _sut_A.TcoSequencerTest := eTcoSequenceTests.StepMode;
            _sut_N.TcoSequencerTest := eTcoSequenceTests.StepMode;
            _sut_A.SetStepMode(); //Set sequencer into the step mode
            _sut_N.SetStepMode(); //Set sequencer into the step mode
            _sut_A.SetSequenceAsChecked(); //Set sequence as checked, so no StepID uniqueness is performed on next sequence execution
            _sut_N.SetSequenceAsChecked(); //Set sequence as checked, so no StepID uniqueness is performed on next sequence execution
            _sut_A.ClearNumberOfSteps();
            _sut_N.ClearNumberOfSteps();
            _sut_A.SetCurrentStep(inStepID := _currentStepId, inStepDescription := _currentStepDescription);
            _sut_N.SetCurrentStep(inStepID := _currentStepId, inStepDescription := _currentStepDescription);
            _sut_A.TotalStepNumber := _totalStepNumber;
            _sut_N.TotalStepNumber := _totalStepNumber;
            _sut_A.SaveNumberOfStepsInSequence();
            _sut_N.SaveNumberOfStepsInSequence();
            _plcCycleCounter := 0;
            _arranged := TRUE;
            RETURN;
        END_IF

        IF NOT _done THEN
            _sut_A.SequenceRun := _plcCycleCounter;
            _sut_N.SequenceRun := _plcCycleCounter;
            _sut_A._RunExecutionSubstitute();
            _sut_N._RunExecutionSubstitute();
            _sut_A.SaveNumberOfStepsInSequence();
            _sut_N.SaveNumberOfStepsInSequence();
        END_IF

        _done := _plcCycleCounter >= _totalStepNumber + 1;
        ProbeDoneWhen(_done);
    {endregion}
    {region "T582_InvalidMode"}
    eTcoSequenceTests.InvalidMode:
        IF NOT _arranged THEN
            _sut_A.TcoSequencerTest := eTcoSequenceTests.SetStepMode;
            _sut_N.TcoSequencerTest := eTcoSequenceTests.SetStepMode;
            _sut_A.SetCyclicMode(); //Set sequencer into the cyclic mode
            _sut_N.SetCyclicMode(); //Set sequencer into the cyclic mode
            _sut_A.SetSequenceAsChecked(); //Set sequence as checked, so no StepID uniqueness is performed on next sequence execution
            _sut_N.SetSequenceAsChecked(); //Set sequence as checked, so no StepID uniqueness is performed on next sequence execution
            _sut_A.SetNumberOfSteps(_totalStepNumber);
            _sut_N.SetNumberOfSteps(_totalStepNumber);
            _sut_A.SetCurrentStep(inStepID := _currentStepId, inStepDescription := _currentStepDescription);
            _sut_N.SetCurrentStep(inStepID := _currentStepId, inStepDescription := _currentStepDescription);
            _sut_A.TotalStepNumber := _totalStepNumber;
            _sut_N.TotalStepNumber := _totalStepNumber;
            _sut_A.SaveNumberOfStepsInSequence();
            _sut_N.SaveNumberOfStepsInSequence();
            _plcCycleCounter := 0;
            _arranged := TRUE;
            RETURN;
        END_IF

        IF NOT _done THEN
            _sut_A.SequenceRun := _plcCycleCounter;
            _sut_N.SequenceRun := _plcCycleCounter;

            IF _plcCycleCounter = 1 THEN
                _sut_A.SequencerOpen();
                _sut_N.SequencerOpen();

                FOR i := 0 TO _totalStepNumber - 1 DO
                    IF _sut_A._Step(i, TRUE, CONCAT('Step ', INT_TO_STRING(i))) THEN
                        _sut_A._StepCompleteWhen(TRUE);
                    END_IF

                    IF _sut_N._Step(i, TRUE, CONCAT('Step ', INT_TO_STRING(i))) THEN
                        _sut_N._StepCompleteWhen(TRUE);
                    END_IF
                END_FOR
            END_IF

            IF _plcCycleCounter = 2 THEN
                _sut_A._Step(_totalStepNumber, TRUE, CONCAT('Step ', INT_TO_STRING(_totalStepNumber)));
                _sut_N._Step(_totalStepNumber, TRUE, CONCAT('Step ', INT_TO_STRING(_totalStepNumber)));
                _sut_A.SequencerClose();
                _sut_N.SequencerClose();
            END_IF

            IF _plcCycleCounter = 3 THEN
                _sut_A.SequencerOpen();
                _sut_N.SequencerOpen();

                FOR i := 0 TO _totalStepNumber DO
                    _sut_A._Step(i, TRUE, CONCAT('Step ', INT_TO_STRING(i)));
                    _sut_N._Step(i, TRUE, CONCAT('Step ', INT_TO_STRING(i)));
                END_FOR

                _sut_A.SequencerClose();
                _sut_N.SequencerClose();
            END_IF

            _sut_A.SaveNumberOfStepsInSequence();
            _sut_N.SaveNumberOfStepsInSequence();
        END_IF

        _done := _plcCycleCounter >= 3;
        ProbeDoneWhen(_done);
    {endregion}
    {region "T582_StepInError"}
    eTcoSequenceTests.StepInError:
        IF NOT _arranged THEN
            _sut_A.TcoSequencerTest := eTcoSequenceTests.StepInError;
            _sut_N.TcoSequencerTest := eTcoSequenceTests.StepInError;
            _sut_A.SetCyclicMode(); //Set sequencer into the cyclic mode
            _sut_N.SetCyclicMode(); //Set sequencer into the cyclic mode
            _sut_A.SetSequenceAsChecked(); //Set sequence as checked, so no StepID uniqueness is performed on next sequence execution
            _sut_N.SetSequenceAsChecked(); //Set sequence as checked, so no StepID uniqueness is performed on next sequence execution
            _sut_A.SetNumberOfSteps(_totalStepNumber);
            _sut_N.SetNumberOfSteps(_totalStepNumber);
            _sut_A.SetCurrentStep(inStepID := _currentStepId, inStepDescription := _currentStepDescription);
            _sut_N.SetCurrentStep(inStepID := _currentStepId, inStepDescription := _currentStepDescription);
            _sut_A.TotalStepNumber := _totalStepNumber;
            _sut_N.TotalStepNumber := _totalStepNumber;
            _sut_A.SaveNumberOfStepsInSequence();
            _sut_N.SaveNumberOfStepsInSequence();
            _plcCycleCounter := 0;
            _arranged := TRUE;
            RETURN;
        END_IF

        IF NOT _done THEN
            _sut_A.SequenceRun := _plcCycleCounter;
            _sut_N.SequenceRun := _plcCycleCounter;

            IF _plcCycleCounter = 1 THEN
                _sut_A.SequencerOpen();
                _sut_N.SequencerOpen();

                FOR i := 0 TO _totalStepNumber - 1 DO
                    IF _sut_A._Step(i, TRUE, CONCAT('Step ', INT_TO_STRING(i))) THEN
                        _sut_A._StepCompleteWhen(TRUE);
                    END_IF

                    IF _sut_N._Step(i, TRUE, CONCAT('Step ', INT_TO_STRING(i))) THEN
                        _sut_N._StepCompleteWhen(TRUE);
                    END_IF
                END_FOR
            END_IF

            IF _plcCycleCounter = 2 THEN
                _sut_A._Step(_totalStepNumber, TRUE, CONCAT('Step ', INT_TO_STRING(_totalStepNumber)));
                _sut_N._Step(_totalStepNumber, TRUE, CONCAT('Step ', INT_TO_STRING(_totalStepNumber)));
                _sut_A.SequencerClose();
                _sut_N.SequencerClose();
            END_IF

            IF _plcCycleCounter = 3 THEN
                _sut_A.SequencerOpen();
                _sut_N.SequencerOpen();

                FOR i := 0 TO _totalStepNumber DO
                    _sut_A._Step(i, TRUE, CONCAT('Step ', INT_TO_STRING(i)));
                    _sut_N._Step(i, TRUE, CONCAT('Step ', INT_TO_STRING(i)));
                END_FOR

                _sut_A.SequencerClose();
                _sut_N.SequencerClose();
            END_IF

            _sut_A.SaveNumberOfStepsInSequence();
            _sut_N.SaveNumberOfStepsInSequence();
        END_IF

        _done := _plcCycleCounter >= 3;
        ProbeDoneWhen(_done);
    {endregion}
    {region "T590_CheckStepIdUniquenessStepMode"}
    eTcoSequenceTests.CheckStepIdUniquenessStepMode:
        IF NOT _arranged THEN
            _sut_A.SetStepMode(); //Set sequencer into the step mode
            _sut_N.SetStepMode(); //Set sequencer into the step mode
            _sut_A.SetSequenceAsNotChecked(); //Set sequence as not checked, so StepId uniqueness is going to be performed on next sequence run
            _sut_N.SetSequenceAsNotChecked(); //Set sequence as not checked, so StepId uniqueness is going to be performed on next sequence run
            _sut_A.ClearNumberOfSteps(); //Clear internal step counters, so number of steps is going to be counted again on next sequence run
            _sut_N.ClearNumberOfSteps(); //Clear internal step counters, so number of steps is going to be counted again on next sequence run
            _sut_A.Enabled := TRUE;
            _sut_A.RunOneStep := FALSE;
            _sut_A.RunAllSteps := TRUE;
            _sut_A.FinishStep := TRUE;
            _sut_A.StepId := _stepId;
            _sut_A.StepDescription := _stepDescription;
            _sut_N.Enabled := TRUE;
            _sut_N.RunOneStep := FALSE;
            _sut_N.RunAllSteps := TRUE;
            _sut_N.FinishStep := TRUE;
            _sut_N.StepId := _stepId;
            _sut_N.StepDescription := _stepDescription;
            _sut_A.SetCurrentStep(inStepID := _currentStepId, inStepDescription := _currentStepDescription);
            _sut_N.SetCurrentStep(inStepID := _currentStepId, inStepDescription := _currentStepDescription);
            _sut_A.TcoSequencerTest := eTcoSequenceTests.CheckStepIdUniquenessStepMode;
            _sut_N.TcoSequencerTest := eTcoSequenceTests.CheckStepIdUniquenessStepMode;
            _sut_A.SaveNumberOfStepsInSequence();
            _sut_N.SaveNumberOfStepsInSequence();
            _plcCycleCounter := 0;
            _arranged := TRUE;
            RETURN;
        END_IF

        IF NOT _done THEN
            IF _plcCycleCounter = 3 THEN
                _sut_A._StepIn();
                _sut_N._StepIn();
            END_IF

            _sut_A._RunExecutionSubstitute();
            _sut_N._RunExecutionSubstitute();

            IF _plcCycleCounter = 4 THEN
                _sut_A.Restore();
                _sut_N.Restore();
            END_IF

            _sut_A.SaveNumberOfStepsInSequence();
            _sut_N.SaveNumberOfStepsInSequence();
        END_IF

        _done := _plcCycleCounter >= 4;

        IF _done THEN
            _sut_A.TcoSequencerTest := eTcoSequenceTests.none;
            _sut_N.TcoSequencerTest := eTcoSequenceTests.none;
        END_IF

        ProbeDoneWhen(_done);
    {endregion}
    {region "T594_NotUniqueStepIdInStepMode"}
    eTcoSequenceTests.NotUniqueStepIdInStepMode:
        IF NOT _arranged THEN
            _sut_A.TcoSequencerTest := eTcoSequenceTests.NotUniqueStepIdInStepMode;
            _sut_N.TcoSequencerTest := eTcoSequenceTests.NotUniqueStepIdInStepMode;
            _sut_A.SetStepMode(); //Set sequencer into the step mode
            _sut_N.SetStepMode(); //Set sequencer into the step mode
            _sut_A.Enabled := TRUE;
            _sut_A.RunOneStep := FALSE;
            _sut_A.RunAllSteps := FALSE;
            _sut_A.FinishStep := TRUE;
            _sut_A.StepId := _stepId;
            _sut_N.Enabled := TRUE;
            _sut_N.RunOneStep := FALSE;
            _sut_N.RunAllSteps := FALSE;
            _sut_N.FinishStep := TRUE;
            _sut_N.StepId := _stepId;
            _sut_A.SetCurrentStep(inStepID := _currentStepId, inStepDescription := _currentStepDescription);
            _sut_N.SetCurrentStep(inStepID := _currentStepId, inStepDescription := _currentStepDescription);
            _sut_A.SaveNumberOfStepsInSequence();
            _sut_N.SaveNumberOfStepsInSequence();
            _plcCycleCounter := 0;
            _arranged := TRUE;
            RETURN;
        END_IF

        IF NOT _done THEN
            IF _plcCycleCounter = 2 THEN
                _Sut_A.RunOneStep := TRUE;
                _Sut_N.RunOneStep := TRUE;
            END_IF

            _sut_A._RunExecutionSubstitute();
            _sut_N._RunExecutionSubstitute();
            _sut_A.SaveNumberOfStepsInSequence();
            _sut_N.SaveNumberOfStepsInSequence();
            _done := _plcCycleCounter >= 2;
        END_IF

        IF _done THEN
            ProbeDoneWhen(_done);
        END_IF
    {endregion}
    {region "T597_AfterErrorResetInStepMode"}
    eTcoSequenceTests.AfterErrorResetInStepMode:
        IF NOT _arranged THEN
            _sut_A.TcoSequencerTest := eTcoSequenceTests.AfterErrorRestore;
            _sut_N.TcoSequencerTest := eTcoSequenceTests.AfterErrorRestore;
            _sut_A.SetStepMode();
            _sut_N.SetStepMode();
            _sut_A.SaveNumberOfStepsInSequence();
            _sut_N.SaveNumberOfStepsInSequence();
            _plcCycleCounter := 0;
            _arranged := TRUE;
            RETURN;
        END_IF

        IF NOT _done THEN
            IF _plcCycleCounter = 3 THEN
                _sut_A._StepIn();
                _sut_N._StepIn();
            END_IF

            _sut_A._RunExecutionSubstitute();
            _sut_N._RunExecutionSubstitute();
            _sut_A.SaveNumberOfStepsInSequence();
            _sut_N.SaveNumberOfStepsInSequence();
            _done := _plcCycleCounter >= 4;
        END_IF

        IF _done THEN
            ProbeDoneWhen(_done);
        END_IF
    {endregion}
    {region "T601_InvalidModeDetailed"}
    eTcoSequenceTests.InvalidModeDetailed:
        IF NOT _arranged THEN
            _sut_A.TcoSequencerTest := eTcoSequenceTests.InvalidModeDetailed;
            _sut_N.TcoSequencerTest := eTcoSequenceTests.InvalidModeDetailed;
            _sut_A.SetSequenceAsNotChecked();
            _sut_N.SetSequenceAsNotChecked();
            _sut_A.ClearNumberOfSteps();
            _sut_N.ClearNumberOfSteps();
            _sut_A.SetCurrentStep(_currentStepId, _currentStepDescription);
            _sut_N.SetCurrentStep(_currentStepId, _currentStepDescription);
            _sut_A.StepId := _stepId;
            _sut_N.StepId := _stepId;
            _sut_A.StepDescription := _stepDescription;
            _sut_N.StepDescription := _stepDescription;
            _sut_A.Enabled := TRUE;
            _sut_N.Enabled := TRUE;
            _sut_A.RunOneStep := FALSE;
            _sut_N.RunOneStep := FALSE;
            _sut_A.RunAllSteps := TRUE;
            _sut_N.RunAllSteps := TRUE;
            _sut_A.FinishStep := TRUE;
            _sut_N.FinishStep := TRUE;
            _sut_A.SetStepMode();
            _sut_N.SetStepMode();
            _sut_A.SaveNumberOfStepsInSequence();
            _sut_N.SaveNumberOfStepsInSequence();
            _plcCycleCounter := 0;
            _arranged := TRUE;
            RETURN;
        END_IF

        IF NOT _done THEN
            IF _plcCycleCounter = 2 THEN
                _sut_A.SetInvalidMode();
                _sut_N.SetInvalidMode();
                _sut_A.RunOneStep := TRUE;
                _sut_N.RunOneStep := TRUE;
                _sut_A.RunAllSteps := FALSE;
                _sut_N.RunAllSteps := FALSE;
            END_IF

            _sut_A._RunExecutionSubstitute();
            _sut_N._RunExecutionSubstitute();
            _sut_A.SaveNumberOfStepsInSequence();
            _sut_N.SaveNumberOfStepsInSequence();
            _done := _plcCycleCounter >= 2;
        END_IF

        IF _done THEN
            ProbeDoneWhen(_done);
        END_IF
    {endregion}
    {region "T604_StepInErrorDetailed"}
    eTcoSequenceTests.StepInErrorDetailed:
        IF NOT _arranged THEN
            _sut_A.TcoSequencerTest := eTcoSequenceTests.StepInErrorDetailed;
            _sut_N.TcoSequencerTest := eTcoSequenceTests.StepInErrorDetailed;
            _sut_A.SetSequenceAsNotChecked();
            _sut_N.SetSequenceAsNotChecked();
            _sut_A.ClearNumberOfSteps();
            _sut_N.ClearNumberOfSteps();
            _sut_A.SetCurrentStep(_currentStepId, _currentStepDescription);
            _sut_N.SetCurrentStep(_currentStepId, _currentStepDescription);
            _sut_A.StepId := _stepId;
            _sut_N.StepId := _stepId;
            _sut_A.StepDescription := _stepDescription;
            _sut_N.StepDescription := _stepDescription;
            _sut_A.Enabled := TRUE;
            _sut_N.Enabled := TRUE;
            _sut_A.RunOneStep := FALSE;
            _sut_N.RunOneStep := FALSE;
            _sut_A.RunAllSteps := TRUE;
            _sut_N.RunAllSteps := TRUE;
            _sut_A.FinishStep := TRUE;
            _sut_N.FinishStep := TRUE;
            _sut_A.SetStepMode();
            _sut_N.SetStepMode();
            _sut_A.SaveNumberOfStepsInSequence();
            _sut_N.SaveNumberOfStepsInSequence();
            _plcCycleCounter := 0;
            _arranged := TRUE;
            RETURN;
        END_IF

        IF NOT _done THEN
            IF _plcCycleCounter = 2 THEN
                _sut_A.SetCurrentStepToErrorState();
                _sut_N.SetCurrentStepToErrorState();
                _sut_A.RunOneStep := TRUE;
                _sut_N.RunOneStep := TRUE;
                _sut_A.RunAllSteps := FALSE;
                _sut_N.RunAllSteps := FALSE;
            END_IF

            _sut_A._RunExecutionSubstitute();
            _sut_N._RunExecutionSubstitute();
            _sut_A.SaveNumberOfStepsInSequence();
            _sut_N.SaveNumberOfStepsInSequence();
            _done := _plcCycleCounter >= 2;
        END_IF

        IF _done THEN
            ProbeDoneWhen(_done);
        END_IF
    {endregion}
    {region "T611_StepModeStepIn"}
    eTcoSequenceTests.StepModeStepIn:
        IF NOT _arranged THEN
            _sut_A.TcoSequencerTest := eTcoSequenceTests.StepModeStepIn;
            _sut_N.TcoSequencerTest := eTcoSequenceTests.StepModeStepIn;
            _sut_A.SetSequenceAsChecked();
            _sut_N.SetSequenceAsChecked();
            _sut_A.SetNumberOfSteps(_totalStepNumber);
            _sut_N.SetNumberOfSteps(_totalStepNumber);
            _sut_A.TotalStepNumber := _totalStepNumber;
            _sut_N.TotalStepNumber := _totalStepNumber;
            _sut_A.SetCurrentStep(_currentStepId, _currentStepDescription);
            _sut_N.SetCurrentStep(_currentStepId, _currentStepDescription);
            _sut_A.StepId := _stepId;
            _sut_N.StepId := _stepId;
            _sut_A.StepDescription := _stepDescription;
            _sut_N.StepDescription := _stepDescription;
            _sut_A.Enabled := TRUE;
            _sut_N.Enabled := TRUE;
            _sut_A.RunOneStep := FALSE;
            _sut_N.RunOneStep := FALSE;
            _sut_A.RunAllSteps := TRUE;
            _sut_N.RunAllSteps := TRUE;
            _sut_A.FinishStep := TRUE;
            _sut_N.FinishStep := TRUE;
            _sut_A.SetStepMode();
            _sut_N.SetStepMode();
            _sut_A.SaveNumberOfStepsInSequence();
            _sut_N.SaveNumberOfStepsInSequence();
            _plcCycleCounter := 0;
            _arranged := TRUE;
            RETURN;
        END_IF

        IF NOT _done THEN
            _sut_A.SequenceRun := _plcCycleCounter;
            _sut_N.SequenceRun := _plcCycleCounter;
            _sut_A._RunExecutionSubstitute();
            _sut_N._RunExecutionSubstitute();
            _sut_A.SaveNumberOfStepsInSequence();
            _sut_N.SaveNumberOfStepsInSequence();
            _done := _plcCycleCounter >= _totalStepNumber + 1;
        END_IF

        IF _done THEN
            ProbeDoneWhen(_done);
        END_IF
    {endregion}
    {region "T612_StepModeChangeStepIdDuringExecution"}
    eTcoSequenceTests.StepModeChangeStepIdDuringExecution:
        IF NOT _done AND _plcCycleCounter <= 2 THEN
            _sut_A.TcoSequencerTest := eTcoSequenceTests.StepModeChangeStepIdDuringExecution;
            _sut_N.TcoSequencerTest := eTcoSequenceTests.StepModeChangeStepIdDuringExecution;
            _sut_A.SequenceRun := _plcCycleCounter;
            _sut_N.SequenceRun := _plcCycleCounter;
            _sut_A._RunExecutionSubstitute();
            _sut_N._RunExecutionSubstitute();
            _sut_A.SaveNumberOfStepsInSequence();
            _sut_N.SaveNumberOfStepsInSequence();
        END_IF

        IF _plcCycleCounter >= 3 THEN
            _sut_A.Restore();
            _sut_N.Restore();
            _sut_A.SetSequenceAsChecked();
            _sut_N.SetSequenceAsChecked();
            _sut_A.SetNumberOfSteps(_totalStepNumber);
            _sut_N.SetNumberOfSteps(_totalStepNumber);
            _sut_A.TotalStepNumber := _totalStepNumber;
            _sut_N.TotalStepNumber := _totalStepNumber;
            _sut_A.SetStepMode();
            _sut_N.SetStepMode();
            _sut_A.SaveNumberOfStepsInSequence();
            _sut_N.SaveNumberOfStepsInSequence();
        END_IF

        _done := _plcCycleCounter >= 3;

        IF _done THEN
            ProbeDoneWhen(_done);
        END_IF
    {endregion}
    {region "T615_StepModeChangeStepOrder"}
    eTcoSequenceTests.StepModeChangeStepOrder:
        IF NOT _arranged THEN
            _sut_A.TcoSequencerTest := eTcoSequenceTests.StepModeChangeStepOrder;
            _sut_N.TcoSequencerTest := eTcoSequenceTests.StepModeChangeStepOrder;
            _sut_A.SetSequenceAsChecked();
            _sut_N.SetSequenceAsChecked();
            _sut_A.SetNumberOfSteps(_totalStepNumber);
            _sut_N.SetNumberOfSteps(_totalStepNumber);
            _sut_A.TotalStepNumber := _totalStepNumber;
            _sut_N.TotalStepNumber := _totalStepNumber;
            _sut_A.SetCurrentStep(_currentStepId, _currentStepDescription);
            _sut_N.SetCurrentStep(_currentStepId, _currentStepDescription);
            _sut_A.StepId := _stepId;
            _sut_N.StepId := _stepId;
            _sut_A.StepDescription := _stepDescription;
            _sut_N.StepDescription := _stepDescription;
            _sut_A.Enabled := TRUE;
            _sut_N.Enabled := TRUE;
            _sut_A.RunOneStep := FALSE;
            _sut_N.RunOneStep := FALSE;
            _sut_A.RunAllSteps := TRUE;
            _sut_N.RunAllSteps := TRUE;
            _sut_A.FinishStep := TRUE;
            _sut_N.FinishStep := TRUE;
            _sut_A.SetStepMode();
            _sut_N.SetStepMode();
            _sut_A.SaveNumberOfStepsInSequence();
            _sut_N.SaveNumberOfStepsInSequence();
            _plcCycleCounter := 0;
            _arranged := TRUE;
            RETURN;
        END_IF

        IF _plcCycleCounter <= _totalStepNumber + 2 THEN
            _sut_A.SequenceRun := _plcCycleCounter;
            _sut_N.SequenceRun := _plcCycleCounter;
            _sut_A._RunExecutionSubstitute();
            _sut_N._RunExecutionSubstitute();
            _sut_A.SaveNumberOfStepsInSequence();
            _sut_N.SaveNumberOfStepsInSequence();
        END_IF

        IF _plcCycleCounter >= _totalStepNumber + 3 THEN
            _sut_A.Restore();
            _sut_N.Restore();
            _sut_A.SetSequenceAsChecked();
            _sut_N.SetSequenceAsChecked();
            _sut_A.SetNumberOfSteps(_totalStepNumber);
            _sut_N.SetNumberOfSteps(_totalStepNumber);
            _sut_A.TotalStepNumber := _totalStepNumber;
            _sut_N.TotalStepNumber := _totalStepNumber;
            _sut_A.SetStepMode();
            _sut_N.SetStepMode();
            _sut_A.SaveNumberOfStepsInSequence();
            _sut_N.SaveNumberOfStepsInSequence();
        END_IF

        _done := _plcCycleCounter >= _totalStepNumber + 3;

        IF _done THEN
            ProbeDoneWhen(_done);
        END_IF
    {endregion}
    {region "T618_StepModeCommentOutPartOfRunningSequencer"}
    eTcoSequenceTests.StepModeCommentOutPartOfRunningSequencer:
        IF NOT _arranged THEN
            _sut_A.TcoSequencerTest := eTcoSequenceTests.StepModeCommentOutPartOfRunningSequencer;
            _sut_N.TcoSequencerTest := eTcoSequenceTests.StepModeCommentOutPartOfRunningSequencer;
            _sut_A.SetStepMode(); //Set sequencer into the step mode
            _sut_N.SetStepMode(); //Set sequencer into the step mode
            _sut_A.SetSequenceAsChecked(); //Set sequence as checked, so no StepID uniqueness is performed on next sequence execution
            _sut_N.SetSequenceAsChecked(); //Set sequence as checked, so no StepID uniqueness is performed on next sequence execution
            _sut_A.ClearNumberOfSteps(); //Clear internal step counters, so number of steps is going to be counted again on next sequence run
            _sut_N.ClearNumberOfSteps(); //Clear internal step counters, so number of steps is going to be counted again on next sequence run
            _sut_A.SetCurrentStep(inStepID := _currentStepId, inStepDescription := _currentStepDescription);
            _sut_N.SetCurrentStep(inStepID := _currentStepId, inStepDescription := _currentStepDescription);
            _sut_A.TotalStepNumber := _totalStepNumber;
            _sut_N.TotalStepNumber := _totalStepNumber;
            _sut_A.SaveNumberOfStepsInSequence();
            _sut_N.SaveNumberOfStepsInSequence();
            _plcCycleCounter := 0;
            _arranged := TRUE;
            RETURN;
        END_IF

        IF NOT _done THEN
            IF _plcCycleCounter = 3 THEN
                _sut_A.Restore();
                _sut_N.Restore();
                _sut_A.SetSequenceAsChecked(); //Set sequence as checked, so no StepID uniqueness is performed on next sequence execution
                _sut_N.SetSequenceAsChecked(); //Set sequence as checked, so no StepID uniqueness is performed on next sequence execution
                _sut_A.ClearNumberOfSteps(); //Clear internal step counters, so number of steps is going to be counted again on next sequence run
                _sut_N.ClearNumberOfSteps(); //Clear internal step counters, so number of steps is going to be counted again on next sequence run
            END_IF

            _sut_A.SequenceRun := _plcCycleCounter;
            _sut_N.SequenceRun := _plcCycleCounter;
            _sut_A._RunExecutionSubstitute();
            _sut_N._RunExecutionSubstitute();
            _sut_A.SaveNumberOfStepsInSequence();
            _sut_N.SaveNumberOfStepsInSequence();
        END_IF

        _done := _plcCycleCounter >= 3;
        ProbeDoneWhen(_done);
    {endregion}
    {region "T621_StepModeUncommentPartOfRunningSequencer"}
    eTcoSequenceTests.StepModeUncommentPartOfRunningSequencer:
        IF NOT _arranged THEN
            _sut_A.TcoSequencerTest := eTcoSequenceTests.StepModeUncommentPartOfRunningSequencer;
            _sut_N.TcoSequencerTest := eTcoSequenceTests.StepModeUncommentPartOfRunningSequencer;
            _sut_A.SetStepMode(); //Set sequencer into the step mode
            _sut_N.SetStepMode(); //Set sequencer into the step mode
            _sut_A.SetSequenceAsChecked(); //Set sequence as checked, so no StepID uniqueness is performed on next sequence execution
            _sut_N.SetSequenceAsChecked(); //Set sequence as checked, so no StepID uniqueness is performed on next sequence execution
            _sut_A.ClearNumberOfSteps(); //Clear internal step counters, so number of steps is going to be counted again on next sequence run
            _sut_N.ClearNumberOfSteps(); //Clear internal step counters, so number of steps is going to be counted again on next sequence run
            _sut_A.SetCurrentStep(inStepID := _currentStepId, inStepDescription := _currentStepDescription);
            _sut_N.SetCurrentStep(inStepID := _currentStepId, inStepDescription := _currentStepDescription);
            _sut_A.TotalStepNumber := _totalStepNumber;
            _sut_N.TotalStepNumber := _totalStepNumber;
            _sut_A.SaveNumberOfStepsInSequence();
            _sut_N.SaveNumberOfStepsInSequence();
            _plcCycleCounter := 0;
            _arranged := TRUE;
            RETURN;
        END_IF

        IF NOT _done THEN
            _sut_A.SequenceRun := _plcCycleCounter;
            _sut_N.SequenceRun := _plcCycleCounter;
            _sut_A._RunExecutionSubstitute();
            _sut_N._RunExecutionSubstitute();
            _sut_A.SaveNumberOfStepsInSequence();
            _sut_N.SaveNumberOfStepsInSequence();
        END_IF

        _done := _plcCycleCounter >= 2;
        ProbeDoneWhen(_done);
    {endregion}
    {region "T631_StepModeRequestStepFromLowerToHigher"}
    eTcoSequenceTests.StepModeRequestStepFromLowerToHigher:
        IF NOT _arranged THEN
            _sut_A.TcoSequencerTest := eTcoSequenceTests.StepModeRequestStepFromLowerToHigher;
            _sut_N.TcoSequencerTest := eTcoSequenceTests.StepModeRequestStepFromLowerToHigher;
            _sut_A.SetStepMode(); //Set sequencer into the step mode
            _sut_N.SetStepMode(); //Set sequencer into the step mode
            _sut_A.SetSequenceAsChecked(); //Set sequence as checked, so no StepID uniqueness is performed on next sequence execution
            _sut_N.SetSequenceAsChecked(); //Set sequence as checked, so no StepID uniqueness is performed on next sequence execution
            _sut_A.ClearNumberOfSteps(); //Clear internal step counters, so number of steps is going to be counted again on next sequence run
            _sut_N.ClearNumberOfSteps(); //Clear internal step counters, so number of steps is going to be counted again on next sequence run
            _sut_A.SetCurrentStep(inStepID := _currentStepId, inStepDescription := _currentStepDescription);
            _sut_N.SetCurrentStep(inStepID := _currentStepId, inStepDescription := _currentStepDescription);
            _sut_A.TotalStepNumber := _totalStepNumber;
            _sut_N.TotalStepNumber := _totalStepNumber;
            _sut_A.ReqStep := _reqStep;
            _sut_N.ReqStep := _reqStep;
            _sut_A.ReqStepNotExists := _reqStepNotExists;
            _sut_N.ReqStepNotExists := _reqStepNotExists;
            _sut_A.SaveNumberOfStepsInSequence();
            _sut_N.SaveNumberOfStepsInSequence();
            _plcCycleCounter := 0;
            _arranged := TRUE;
            RETURN;
        END_IF

        IF NOT _done THEN
            _sut_A.SequenceRun := _plcCycleCounter;
            _sut_N.SequenceRun := _plcCycleCounter;
            _sut_A._RunExecutionSubstitute();
            _sut_N._RunExecutionSubstitute();
            _sut_A.SaveNumberOfStepsInSequence();
            _sut_N.SaveNumberOfStepsInSequence();
        END_IF

        _done := _plcCycleCounter >= 2;
        ProbeDoneWhen(_done);
    {endregion}
    {region "T633_StepModeRequestStepFromHigherToLower"}
    eTcoSequenceTests.StepModeRequestStepFromHigherToLower:
        IF NOT _arranged THEN
            _sut_A.TcoSequencerTest := eTcoSequenceTests.StepModeRequestStepFromHigherToLower;
            _sut_N.TcoSequencerTest := eTcoSequenceTests.StepModeRequestStepFromHigherToLower;
            _sut_A.SetStepMode(); //Set sequencer into the step mode
            _sut_N.SetStepMode(); //Set sequencer into the step mode
            _sut_A.SetSequenceAsChecked(); //Set sequence as checked, so no StepID uniqueness is performed on next sequence execution
            _sut_N.SetSequenceAsChecked(); //Set sequence as checked, so no StepID uniqueness is performed on next sequence execution
            _sut_A.SetNumberOfSteps(_totalStepNumber);
            _sut_N.SetNumberOfSteps(_totalStepNumber);
            _sut_A.SetCurrentStep(inStepID := _currentStepId, inStepDescription := _currentStepDescription);
            _sut_N.SetCurrentStep(inStepID := _currentStepId, inStepDescription := _currentStepDescription);
            _sut_A.TotalStepNumber := _totalStepNumber;
            _sut_N.TotalStepNumber := _totalStepNumber;
            _sut_A.ReqStep := _reqStep;
            _sut_N.ReqStep := _reqStep;
            _sut_A.ReqStepNotExists := _reqStepNotExists;
            _sut_N.ReqStepNotExists := _reqStepNotExists;
            _sut_A.SaveNumberOfStepsInSequence();
            _sut_N.SaveNumberOfStepsInSequence();
            _plcCycleCounter := 0;
            _arranged := TRUE;
            RETURN;
        END_IF

        IF NOT _done THEN
            _sut_A.SequenceRun := _plcCycleCounter;
            _sut_N.SequenceRun := _plcCycleCounter;
            _sut_A._RunExecutionSubstitute();
            _sut_N._RunExecutionSubstitute();
            _sut_A.SaveNumberOfStepsInSequence();
            _sut_N.SaveNumberOfStepsInSequence();
        END_IF

        _done := _plcCycleCounter >= _reqStep + 7;
        ProbeDoneWhen(_done);
    {endregion}
    {region "T635_StepModeRequestStepToNotExistingStep"}
    eTcoSequenceTests.StepModeRequestStepToNotExistingStep:
        IF NOT _arranged THEN
            _sut_A.TcoSequencerTest := eTcoSequenceTests.RequestStepToNotExistingStep;
            _sut_N.TcoSequencerTest := eTcoSequenceTests.RequestStepToNotExistingStep;
            _sut_A.SetStepMode(); //Set sequencer into the step mode
            _sut_N.SetStepMode(); //Set sequencer into the step mode
            _sut_A.SetSequenceAsChecked(); //Set sequence as checked, so no StepID uniqueness is performed on next sequence execution
            _sut_N.SetSequenceAsChecked(); //Set sequence as checked, so no StepID uniqueness is performed on next sequence execution
            _sut_A.SetNumberOfSteps(_totalStepNumber);
            _sut_N.SetNumberOfSteps(_totalStepNumber);
            _sut_A.SetCurrentStep(inStepID := _currentStepId, inStepDescription := _currentStepDescription);
            _sut_N.SetCurrentStep(inStepID := _currentStepId, inStepDescription := _currentStepDescription);
            _sut_A.TotalStepNumber := _totalStepNumber;
            _sut_N.TotalStepNumber := _totalStepNumber;
            _sut_A.ReqStep := _reqStep;
            _sut_N.ReqStep := _reqStep;
            _sut_A.ReqStepNotExists := _reqStepNotExists;
            _sut_N.ReqStepNotExists := _reqStepNotExists;
            _sut_A.SaveNumberOfStepsInSequence();
            _sut_N.SaveNumberOfStepsInSequence();
            _plcCycleCounter := 0;
            _arranged := TRUE;
            RETURN;
        END_IF

        IF _plcCycleCounter = 4 THEN
            _sut_A.Restore();
            _sut_N.Restore();
            _sut_A.SetStepMode(); //Set sequencer into the step mode
            _sut_N.SetStepMode(); //Set sequencer into the step mode
            _sut_A.SetSequenceAsChecked(); //Set sequence as checked, so no StepID uniqueness is performed on next sequence execution
            _sut_N.SetSequenceAsChecked(); //Set sequence as checked, so no StepID uniqueness is performed on next sequence execution
            _sut_A.SetNumberOfSteps(_totalStepNumber);
            _sut_N.SetNumberOfSteps(_totalStepNumber);
            _sut_A.SetCurrentStep(inStepID := _currentStepId, inStepDescription := _currentStepDescription);
            _sut_N.SetCurrentStep(inStepID := _currentStepId, inStepDescription := _currentStepDescription);
            _sut_A.TotalStepNumber := _totalStepNumber;
            _sut_N.TotalStepNumber := _totalStepNumber;
        END_IF

        IF NOT _done THEN
            _sut_A.SequenceRun := _plcCycleCounter;
            _sut_N.SequenceRun := _plcCycleCounter;
            _sut_A._RunExecutionSubstitute();
            _sut_N._RunExecutionSubstitute();
            _sut_A.SaveNumberOfStepsInSequence();
            _sut_N.SaveNumberOfStepsInSequence();
        END_IF

        _done := _plcCycleCounter >= 4;
        ProbeDoneWhen(_done);
    {endregion}
    {region "T640_StepModeRequestStepWhilePreviousRequestStepHasnotBeenYetProcessed"}
    eTcoSequenceTests.StepModeRequestStepWhilePreviousRequestStepHasnotBeenYetProcessed:
        IF NOT _arranged THEN
            _sut_A.TcoSequencerTest := eTcoSequenceTests.StepModeRequestStepWhilePreviousRequestStepHasnotBeenYetProcessed;
            _sut_N.TcoSequencerTest := eTcoSequenceTests.StepModeRequestStepWhilePreviousRequestStepHasnotBeenYetProcessed;
            _sut_A.SetStepMode(); //Set sequencer into the step mode
            _sut_N.SetStepMode(); //Set sequencer into the step mode
            _sut_A.SetSequenceAsChecked(); //Set sequence as checked, so no StepID uniqueness is performed on next sequence execution
            _sut_N.SetSequenceAsChecked(); //Set sequence as checked, so no StepID uniqueness is performed on next sequence execution
            _sut_A.SetNumberOfSteps(_totalStepNumber);
            _sut_N.SetNumberOfSteps(_totalStepNumber);
            _sut_A.SetCurrentStep(inStepID := _currentStepId, inStepDescription := _currentStepDescription);
            _sut_N.SetCurrentStep(inStepID := _currentStepId, inStepDescription := _currentStepDescription);
            _sut_A.TotalStepNumber := _totalStepNumber;
            _sut_N.TotalStepNumber := _totalStepNumber;
            _sut_A.ReqStep := _reqStep;
            _sut_N.ReqStep := _reqStep;
            _sut_A.ReqStepNotExists := _reqStepNotExists;
            _sut_N.ReqStepNotExists := _reqStepNotExists;
            _sut_A.SaveNumberOfStepsInSequence();
            _sut_N.SaveNumberOfStepsInSequence();
            _plcCycleCounter := 0;
            _arranged := TRUE;
            RETURN;
        END_IF

        IF NOT _done THEN
            _sut_A.SequenceRun := _plcCycleCounter;
            _sut_N.SequenceRun := _plcCycleCounter;
            _sut_A._RunExecutionSubstitute();
            _sut_N._RunExecutionSubstitute();
            _sut_A.SaveNumberOfStepsInSequence();
            _sut_N.SaveNumberOfStepsInSequence();
        END_IF

        _done := TRUE;
        ProbeDoneWhen(_done);
    {endregion}
    {region "T641_StepModeDisabledStep"}
    eTcoSequenceTests.StepModeDisabledStep:
        IF NOT _arranged THEN
            _sut_A.TcoSequencerTest := eTcoSequenceTests.StepModeDisabledStep;
            _sut_N.TcoSequencerTest := eTcoSequenceTests.StepModeDisabledStep;
            _sut_A.SetStepMode(); //Set sequencer into the step mode
            _sut_N.SetStepMode(); //Set sequencer into the step mode
            _sut_A.SetSequenceAsChecked(); //Set sequence as checked, so no StepID uniqueness is performed on next sequence execution
            _sut_N.SetSequenceAsChecked(); //Set sequence as checked, so no StepID uniqueness is performed on next sequence execution
            _sut_A.SetNumberOfSteps(_totalStepNumber);
            _sut_N.SetNumberOfSteps(_totalStepNumber);
            _sut_A.TotalStepNumber := _totalStepNumber;
            _sut_N.TotalStepNumber := _totalStepNumber;
            _sut_A.SaveNumberOfStepsInSequence();
            _sut_N.SaveNumberOfStepsInSequence();
            _plcCycleCounter := 0;
            _arranged := TRUE;
            RETURN;
        END_IF

        IF NOT _done THEN
            _sut_A.SequenceRun := _plcCycleCounter;
            _sut_N.SequenceRun := _plcCycleCounter;
            _sut_A._RunExecutionSubstitute();
            _sut_N._RunExecutionSubstitute();
            _sut_A.SaveNumberOfStepsInSequence();
            _sut_N.SaveNumberOfStepsInSequence();
        END_IF

        _done := _plcCycleCounter >= 6;
        ProbeDoneWhen(_done);
    {endregion}
    {region "T670_StepModeStepForwardBackward"}
    eTcoSequenceTests.StepModeStepForwardBackward:
        IF NOT _arranged THEN
            _sut_A.TcoSequencerTest := eTcoSequenceTests.StepModeStepForwardBackward;
            _sut_N.TcoSequencerTest := eTcoSequenceTests.StepModeStepForwardBackward;
            _sut_A.SetStepMode(); //Set sequencer into the step mode
            _sut_N.SetStepMode(); //Set sequencer into the step mode
            _sut_A.SetSequenceAsChecked(); //Set sequence as checked, so no StepID uniqueness is performed on next sequence execution
            _sut_N.SetSequenceAsChecked(); //Set sequence as checked, so no StepID uniqueness is performed on next sequence execution
            _sut_A.SetNumberOfSteps(_totalStepNumber);
            _sut_N.SetNumberOfSteps(_totalStepNumber);
            _sut_A.TotalStepNumber := _totalStepNumber;
            _sut_N.TotalStepNumber := _totalStepNumber;
            _sut_A.SaveNumberOfStepsInSequence();
            _sut_N.SaveNumberOfStepsInSequence();
            _plcCycleCounter := 0;
            _arranged := TRUE;
            RETURN;
        END_IF

        IF NOT _done THEN
            _sut_A.SequenceRun := _plcCycleCounter;
            _sut_N.SequenceRun := _plcCycleCounter;
            _sut_A._RunExecutionSubstitute();
            _sut_N._RunExecutionSubstitute();
            _sut_A.SaveNumberOfStepsInSequence();
            _sut_N.SaveNumberOfStepsInSequence();
        END_IF

        _done := _plcCycleCounter >= 9;
        ProbeDoneWhen(_done);
    {endregion}
    {region "T681_StepModeStepInDetailed"}
    eTcoSequenceTests.StepModeStepInDetailed:
        IF NOT _arranged THEN
            _sut_A.TcoSequencerTest := eTcoSequenceTests.StepModeStepInDetailed;
            _sut_N.TcoSequencerTest := eTcoSequenceTests.StepModeStepInDetailed;
            _sut_A.SetStepMode(); //Set sequencer into the step mode
            _sut_N.SetStepMode(); //Set sequencer into the step mode
            _sut_A.SetSequenceAsChecked(); //Set sequence as checked, so no StepID uniqueness is performed on next sequence execution
            _sut_N.SetSequenceAsChecked(); //Set sequence as checked, so no StepID uniqueness is performed on next sequence execution
            _sut_A.SetNumberOfSteps(_totalStepNumber);
            _sut_N.SetNumberOfSteps(_totalStepNumber);
            _sut_A.TotalStepNumber := _totalStepNumber;
            _sut_N.TotalStepNumber := _totalStepNumber;
            _sut_A.SaveNumberOfStepsInSequence();
            _sut_N.SaveNumberOfStepsInSequence();
            _plcCycleCounter := 0;
            _arranged := TRUE;
            RETURN;
        END_IF

        IF NOT _done THEN
            _sut_A.SequenceRun := _plcCycleCounter;
            _sut_N.SequenceRun := _plcCycleCounter;
            _sut_A._RunExecutionSubstitute();
            _sut_N._RunExecutionSubstitute();
            _sut_A.SaveNumberOfStepsInSequence();
            _sut_N.SaveNumberOfStepsInSequence();
        END_IF

        _done := _plcCycleCounter >= 5;
        ProbeDoneWhen(_done);		 
    {region "T691_SwitchStepModeOnDuringStepExecution"}
    eTcoSequenceTests.SwitchStepModeOnDuringStepExecution:
        IF NOT _arranged THEN
            _sut_A.TcoSequencerTest := eTcoSequenceTests.SwitchStepModeOnDuringStepExecution;
            _sut_N.TcoSequencerTest := eTcoSequenceTests.SwitchStepModeOnDuringStepExecution;
            _sut_A.SetCyclicMode(); //Set sequencer into the cyclic mode
            _sut_N.SetCyclicMode(); //Set sequencer into the cyclic mode
            _sut_A.SetSequenceAsChecked(); //Set sequence as checked, so no StepID uniqueness is performed on next sequence execution
            _sut_N.SetSequenceAsChecked(); //Set sequence as checked, so no StepID uniqueness is performed on next sequence execution
            _sut_A.SetNumberOfSteps(_totalStepNumber);
            _sut_N.SetNumberOfSteps(_totalStepNumber);
            _sut_A.TotalStepNumber := _totalStepNumber;
            _sut_N.TotalStepNumber := _totalStepNumber;
            _sut_A.SaveNumberOfStepsInSequence();
            _sut_N.SaveNumberOfStepsInSequence();
            _plcCycleCounter := 0;
            _arranged := TRUE;
            RETURN;
        END_IF

        IF NOT _done THEN
            _sut_A.SequenceRun := _plcCycleCounter;
            _sut_N.SequenceRun := _plcCycleCounter;
            _sut_A._RunExecutionSubstitute();
            _sut_N._RunExecutionSubstitute();
            _sut_A.SaveNumberOfStepsInSequence();
            _sut_N.SaveNumberOfStepsInSequence();
        END_IF

        _done := _plcCycleCounter >= 10;
        ProbeDoneWhen(_done);
    {endregion}
    {region "T693_SwitchStepModeStepForwardFromRunningStep"}
    eTcoSequenceTests.StepModeStepForwardFromRunningStep:
        _sut_A.TcoSequencerTest := eTcoSequenceTests.StepModeStepForwardFromRunningStep;
        _sut_N.TcoSequencerTest := eTcoSequenceTests.StepModeStepForwardFromRunningStep;

        IF NOT _done THEN
            _sut_A.SequenceRun := _plcCycleCounter;
            _sut_N.SequenceRun := _plcCycleCounter;
            _sut_A._RunExecutionSubstitute();
            _sut_N._RunExecutionSubstitute();
            _sut_A.SaveNumberOfStepsInSequence();
            _sut_N.SaveNumberOfStepsInSequence();
        END_IF

        _done := _plcCycleCounter >= 20;
        ProbeDoneWhen(_done);
    {endregion}
    {region "T695_SwitchStepModeStepBackwardFromRunningStep"}
    eTcoSequenceTests.StepModeStepBackwardFromRunningStep:
        _sut_A.TcoSequencerTest := eTcoSequenceTests.StepModeStepBackwardFromRunningStep;
        _sut_N.TcoSequencerTest := eTcoSequenceTests.StepModeStepBackwardFromRunningStep;

        IF NOT _done THEN
            _sut_A.SequenceRun := _plcCycleCounter;
            _sut_N.SequenceRun := _plcCycleCounter;
            _sut_A._RunExecutionSubstitute();
            _sut_N._RunExecutionSubstitute();
            _sut_A.SaveNumberOfStepsInSequence();
            _sut_N.SaveNumberOfStepsInSequence();
        END_IF

        _done := _plcCycleCounter >= 20;
        ProbeDoneWhen(_done);
    {endregion}
    {region "T696_SwitchStepModeStepOffFromReadyToRun"}
    eTcoSequenceTests.SwitchStepModeStepOffFromReadyToRun:
        _sut_A.TcoSequencerTest := eTcoSequenceTests.SwitchStepModeStepOffFromReadyToRun;
        _sut_N.TcoSequencerTest := eTcoSequenceTests.SwitchStepModeStepOffFromReadyToRun;

        IF NOT _done THEN
            _sut_A.SequenceRun := _plcCycleCounter;
            _sut_N.SequenceRun := _plcCycleCounter;
            _sut_A._RunExecutionSubstitute();
            _sut_N._RunExecutionSubstitute();
            _sut_A.SaveNumberOfStepsInSequence();
            _sut_N.SaveNumberOfStepsInSequence();
        END_IF

        _done := _plcCycleCounter >= 10;
        ProbeDoneWhen(_done);
    {endregion}
    {region "T697_SwitchStepModeStepOnFromRunning"}
    eTcoSequenceTests.SwitchStepModeStepOnFromRunning:
        _sut_A.TcoSequencerTest := eTcoSequenceTests.SwitchStepModeStepOnFromRunning;
        _sut_N.TcoSequencerTest := eTcoSequenceTests.SwitchStepModeStepOnFromRunning;

        IF NOT _done THEN
            _sut_A.SequenceRun := _plcCycleCounter;
            _sut_N.SequenceRun := _plcCycleCounter;
            _sut_A._RunExecutionSubstitute();
            _sut_N._RunExecutionSubstitute();
            _sut_A.SaveNumberOfStepsInSequence();
            _sut_N.SaveNumberOfStepsInSequence();
        END_IF

        _done := _plcCycleCounter >= 10;
        ProbeDoneWhen(_done);
    {endregion}
    {region "T698_SwitchStepModeStepOffFromRunning"}
    eTcoSequenceTests.SwitchStepModeStepOffFromRunning:
        _sut_A.TcoSequencerTest := eTcoSequenceTests.SwitchStepModeStepOffFromRunning;
        _sut_N.TcoSequencerTest := eTcoSequenceTests.SwitchStepModeStepOffFromRunning;

        IF NOT _done THEN
            _sut_A.SequenceRun := _plcCycleCounter;
            _sut_N.SequenceRun := _plcCycleCounter;
            _sut_A._RunExecutionSubstitute();
            _sut_N._RunExecutionSubstitute();
            _sut_A.SaveNumberOfStepsInSequence();
            _sut_N.SaveNumberOfStepsInSequence();
        END_IF

        _done := _plcCycleCounter >= 10;
        ProbeDoneWhen(_done);
    {endregion}
    {region "T699_OnStateChangeWhenChangingModes"}
    eTcoSequenceTests.OnStateChangeWhenChangingModes:
        IF NOT _arranged THEN
            _sut_A.TcoSequencerTest := eTcoSequenceTests.OnStateChangeWhenChangingModes;
            _sut_N.TcoSequencerTest := eTcoSequenceTests.OnStateChangeWhenChangingModes;
            _sut_A.SetCyclicMode(); //Set sequencer into the cyclic mode
            _sut_N.SetCyclicMode(); //Set sequencer into the cyclic mode
            _sut_A.SetSequenceAsChecked(); //Set sequence as checked, so no StepID uniqueness is performed on next sequence execution
            _sut_N.SetSequenceAsChecked(); //Set sequence as checked, so no StepID uniqueness is performed on next sequence execution
            _sut_A.SetNumberOfSteps(_totalStepNumber);
            _sut_N.SetNumberOfSteps(_totalStepNumber);
            _sut_A.TotalStepNumber := _totalStepNumber;
            _sut_N.TotalStepNumber := _totalStepNumber;
            _sut_A.SaveNumberOfStepsInSequence();
            _sut_N.SaveNumberOfStepsInSequence();
            _sut_A.CyclicCycles := _cyclicCycles;
            _sut_N.CyclicCycles := _cyclicCycles;
            _sut_A.StepInEvents := _stepInEvents;
            _sut_N.StepInEvents := _stepInEvents;
            _sut_A.SequenceCycles := 0;
            _sut_N.SequenceCycles := 0;
            _plcCycleCounter := 0;
            _arranged := TRUE;
            RETURN;
        END_IF

        IF NOT _done THEN
            _sut_A.SequenceRun := _plcCycleCounter;
            _sut_N.SequenceRun := _plcCycleCounter;
            _sut_A._RunExecutionSubstitute();
            _sut_N._RunExecutionSubstitute();
            _sut_A.SaveNumberOfStepsInSequence();
            _sut_N.SaveNumberOfStepsInSequence();
        END_IF

        _done := _plcCycleCounter >= 2 * _cyclicCycles + _stepInEvents + 1;
        ProbeDoneWhen(_done);
{endregion}
	 eTcoSequenceTests.MissedSequenceOpening:
	    _sut_A.Restore();
	 	THIS^._Open();
	 	_sut_A.Step(10, TRUE, '');
		THIS^._Close();
		THIS^.ProbeDoneWhen(TRUE);
	 eTcoSequenceTests.MissedSequenceClosing:
	 	_sut_A.Restore();
	 	THIS^._Open();
	    _sut_A.Open();
	 	_sut_A.Step(10, TRUE, '');
		THIS^._Close();
		_sut_A.Messenger.Clear();
		THIS^._Open();
		 _sut_A.Open();
		_sut_A.Step(10, TRUE, '');
		THIS^.ProbeDoneWhen(TRUE);
	eTcoSequenceTests.FreshStateEntry:
		
		THIS^._sut_A.Open();
		IF(_sut_A.Step(10, TRUE, 'ENTER AND LEAVE')) THEN
			THIS^.FreshStateEntry_enter_and_leave_must_be_true := _sut_A.IsFreshState;
			_sut_A.CompleteStep(); 			 
		END_IF;
		
		IF(_sut_A.Step(20, TRUE, 'ENTER MULTIPLE CYCLES')) THEN 
			IF(FreshStateEntry_counter = 0) THEN
				THIS^.FreshStateEntry_enter_and_two_cycles_on_first_must_be_true := _sut_A.IsFreshState;
			END_IF;				
			THIS^.FreshStateEntry_enter_and_two_cycles_on_second_must_be_false := _sut_A.IsFreshState;
			_sut_A.StepCompleteWhen(FreshStateEntry_counter = 1);
			FreshStateEntry_counter := FreshStateEntry_counter + 1;
		END_IF;
		
		IF(_sut_A.Step(40, TRUE, 'ENTER MULTIPLE CYCLES')) THEN 						
			FreshStateEntry_on_multiple_calls_but_not_first_must_be_false := _sut_A.IsFreshState;											
			FreshStateEntry_counter := FreshStateEntry_counter + 1;
			_sut_A.StepCompleteWhen(FreshStateEntry_counter = 100);
		END_IF;
		
		IF(_sut_A.Step(50, TRUE, 'ENTER MULTIPLE CYCLES')) THEN
			FreshStateEntry_on_request_step_single_call_must_be_true :=	_sut_A.IsFreshState;		 			
			_sut_A.CompleteStep();
			IF(FreshStateEntry_counter = 0) THEN
				_sut_A.RequestStep(70);
			END_IF
		END_IF;
		
		IF(_sut_A.Step(60, TRUE, 'ENTER MULTIPLE CYCLES')) THEN					 			
			_sut_A.RequestStep(50);
			FreshStateEntry_counter := 0;
		END_IF;
		
		IF(_sut_A.Step(70, TRUE, 'ENTER MULTIPLE CYCLES')) THEN					 			
			THIS^.ProbeDoneWhen(TRUE);
		END_IF;
		
		THIS^._sut_A.Close();
END_CASE
END_METHOD

METHOD INTERNAL ReadOutCycleCounters
_startCycles		:=		THIS^.StartCycleCount;
_endCycles			:=		THIS^.EndCycleCount;

_myIdentity			:= 		THIS^.Identity;
END_METHOD

END_FUNCTION_BLOCK

// ---- Tests/TcoSequence/PlcExecuted/TcoSequenceTestType.TcPOU
FUNCTION_BLOCK TcoSequenceTestType EXTENDS TcoCore._internals_TcoSequence
VAR
	_runOneStep							:	BOOL;
	_runAllSteps						:	BOOL;
	_finishStep							:	BOOL;
	_stepId								:	INT;
	_enabled							:	BOOL;
	_stepDescription					:	STRING(254);	
	_currentStepId						:	INT;
	_currentStepDescription				:	STRING(254);
	_myTcoChildState					: 	TcoSequencerTestChildState(THIS^, eRestoreMode.None);
	_onCompleteStepCount 				: 	INT;
	_onSequenceCompleteCount 			: 	INT;
	_onSequencerErrorCount	 			: 	ULINT;
	_onStateChangeCount 				:	ULINT;
	_stateChangeFrom					:	INT;
	_stateChangeTo						:	INT;
	_callRestoreInOnStateChange			:	BOOL;

	_numberOfSteps						:	UINT;
	_previousNumberOfSteps						:	UINT;
	_tcoSequenceTest : eTcoSequenceTests;
    _totalStepNumber : UINT;
	_sequenceRun : ULINT;
	_reqStep : INT;
    _reqStepNotExists : INT;
	_initReqStepCycle		:	UINT;
	
	_postOpenRequestStepCycle : UINT;
	_preCloseRequestStepCycle : UINT;

	_restoreCycleCount : UINT;
	_cyclicCycles :	UINT;
    _stepInEvents :	UINT;
	_sequenceCycles :	UINT;

END_VAR

METHOD _RequestStep
VAR_INPUT
	inRequestedStepId : INT;
END_VAR
THIS^.RequestStep(inRequestedStepId);
END_METHOD

METHOD _RunExecutionSubstitute
VAR_INPUT
END_VAR
THIS^.Open();
THIS^.Main();
THIS^.Close();
END_METHOD

METHOD _SequenceComplete
THIS^.CompleteSequence();
END_METHOD

METHOD INTERNAL _Step : BOOL
VAR_INPUT
	inStepId			:	INT;
	inEnabled			:	BOOL;
	inStepDescription	:	STRING(254);		
END_VAR
_Step := SUPER^.Step(inStepID := inStepId, inEnabled := inEnabled, inStepDescription := inStepDescription);
END_METHOD

METHOD _StepBackward
THIS^.ModeController.StepBackward();
END_METHOD

METHOD _StepCompleteWhen 
VAR_INPUT
	inCondition : BOOL;
END_VAR
THIS^.StepCompleteWhen(inCondition);
END_METHOD

METHOD _StepForward
THIS^.ModeController.StepForward();
END_METHOD

METHOD INTERNAL _StepIn
THIS^.ModeController.StepIn();
END_METHOD

PROPERTY CallRestoreInOnStateChange : BOOL
GET
CallRestoreInOnStateChange := _callRestoreInOnStateChange;
END_GET
SET
_callRestoreInOnStateChange:=CallRestoreInOnStateChange;
END_SET
END_PROPERTY

{attribute 'TcRpcEnable'}
METHOD INTERNAL ChildHasAutoRestoreEnabled : BOOL
ChildHasAutoRestoreEnabled := THIS^._myTcoChildState.IsAutoRestoreEnabled;
END_METHOD

{attribute 'TcRpcEnable'}
METHOD INTERNAL ChildIsAutoRestorable : BOOL
ChildIsAutoRestorable := THIS^._myTcoChildState.AutoRestorable;
END_METHOD

METHOD INTERNAL ClearNumberOfSteps
_stepCounter := 0;
_numberOfStepsInSequence := 0;
_previousNumberOfStepsInSequence := 0;
END_METHOD

PROPERTY CyclicCycles : UINT
GET
CyclicCycles := _cyclicCycles;
END_GET
SET
_cyclicCycles := CyclicCycles;
END_SET
END_PROPERTY

PROPERTY Enabled : BOOL
GET
Enabled := _enabled;
END_GET
SET
_enabled := Enabled;
END_SET
END_PROPERTY

PROPERTY FinishStep : BOOL
GET
FinishStep := _finishStep;
END_GET
SET
_finishStep := FinishStep;
END_SET
END_PROPERTY

{attribute 'TcRpcEnable'}
METHOD INTERNAL GetChildState :	INT
GetChildState := THIS^._myTcoChildState.State;
END_METHOD

{attribute 'TcRpcEnable'}
METHOD GetOrderOfTheCurrentlyEvaluatedStep : UINT
GetOrderOfTheCurrentlyEvaluatedStep := _theOrderOfTheCurrentlyEvaluatedStep;
END_METHOD

{attribute 'TcRpcEnable'}
METHOD GetOrderOfTheCurrentlyExecutedStep : UINT
GetOrderOfTheCurrentlyExecutedStep := _theOrderOfTheCurrentlyExecutedStep;
END_METHOD

{attribute 'TcRpcEnable'}
METHOD GetRequestStepCycle : UINT
GetRequestStepCycle := RequestStepCycle;
END_METHOD

{attribute 'TcRpcEnable'}
METHOD INTERNAL HasAutoRestoreEnabled : BOOL
HasAutoRestoreEnabled := SUPER^.IsAutoRestoreEnabled;
END_METHOD

PROPERTY InitReqStepCycle : UINT
GET
_initReqStepCycle := RequestStepCycle;
InitReqStepCycle:=_initReqStepCycle;
END_GET
SET
_initReqStepCycle:=InitReqStepCycle;
RequestStepCycle := _initReqStepCycle;
END_SET
END_PROPERTY

{attribute 'TcRpcEnable'}
METHOD INTERNAL IsAutoRestorable : BOOL
IsAutoRestorable := SUPER^.AutoRestorable;
END_METHOD

